(* IEC 61131-3 sources: daoli-st-library/DL_MathData (part 20) *)

(* ---- FC_DL_PeriodJitterCalc.st ---- *)
(*
  Name        : FC_DL_PeriodJitterCalc
  Category    : DL_MathData
  Version     : 1.0.0
  Purpose     : 周期序列抖动统计（双精度数组）：均值、样本标准差（n-1 分母）、峰峰抖动（max-min）；/ Period-sequence jitter statistics over a double-precision array: mean, sample standard deviation (n-1) and peak-to-peak jitter (max-min)
  溯源        : 借 t2-1-lgf-math 的分类/参数域组织，clean-room 实现
  Boundary    : ① 计数域钳位：nCount 钳 0..64（容量常量），少于 2 个有效样本时 bValid = FALSE（样本标准差无定义），返回 0.0 哨兵；
                ② 入口有限性闸：任一被统计元素 NaN（x = x 自反）或 Inf（(x-x) = (x-x) 差判）→ 整体 bValid = FALSE（不静默跳过，防抖动被低估）；
                ③ 除零前置：均值除子为常量 1000 换算与 nCount（>= 2 已闸），标准差除子 nCount-1（>= 1 已闸）；
                ④ 数组下标游标 1..nCount 有界遍历（下标全量钳位），不越容量域；
                ⑤ 返回值 = 峰峰抖动 [s]，bValid = FALSE 时不得使用返回值（上层契约）。
*)
FUNCTION FC_DL_PeriodJitterCalc : LREAL
VAR_INPUT
    afPeriods : ARRAY[1..64] OF LREAL;       (* 周期样本数组（连续周期测量值）[s] / Period samples array *)
    nCount    : INT;                         (* 有效样本数，域 0..64（越域钳位）[个] / Valid sample count, clamped *)
END_VAR
VAR_OUTPUT
    fMean     : LREAL;                       (* 周期均值 [s] / Mean period *)
    fStdDev   : LREAL;                       (* 样本标准差（n-1 分母）[s] / Sample standard deviation *)
    bValid    : BOOL;                        (* 结果有效标志（FALSE 时返回值为哨兵零点）[-] / Result validity flag *)
END_VAR
VAR CONSTANT
    DL_PJC_NMAX  : INT   := 64;              (* 数组容量上限（与形参数组域一致）[个] / Array capacity *)
    DL_PJC_NMIN  : INT   := 2;               (* 样本数下限（标准差最少两点）[个] / Sample lower bound *)
    DL_PJC_EPS   : LREAL := 1.0E-12;         (* 双精度判零容差 [s] / Double-precision epsilon *)
    DL_PJC_ONE   : LREAL := 1.0;             (* 游标递进常量 [-] / Cursor step constant *)
END_VAR
VAR
    _nEff  : INT;                            (* 钳位后生效样本数 [个] / Effective sample count *)
    _nIdx  : INT;                            (* 统计游标（每趟重置，R227）[-] / Stats cursor *)
    _fSum  : LREAL;                          (* Σx 中间量 [s] / Sum intermediate *)
    _fMeanI: LREAL;                          (* 均值中间量 [s] / Mean intermediate *)
    _fVar  : LREAL;                          (* Σ(x-x̄)² 中间量 [s²] / Squared-deviation sum *)
    _fStdI : LREAL;                          (* 标准差中间量 [s] / Std intermediate *)
    _fMin  : LREAL;                          (* 样本最小值 [s] / Sample minimum *)
    _fMax  : LREAL;                          (* 样本最大值 [s] / Sample maximum *)
    _bFin  : BOOL;                           (* 全体样本有限性当拍量 / Joint sample finiteness *)
END_VAR

(* —— 段 0：计数域钳位 + 有限性预置 —— *)
bValid := TRUE;                                                                (* 有效标志预置（任一闸命中即翻 FALSE） / Validity preset *)
_nEff := nCount;                                                               (* 生效样本数初值 / Effective count init *)
IF _nEff < 0 THEN
    _nEff := 0;                                                                (* 计数下限钳 0 / Lower clamp *)
END_IF
IF _nEff > DL_PJC_NMAX THEN
    _nEff := DL_PJC_NMAX;                                                      (* 计数上限钳容量（下标全量钳位） / Upper clamp to capacity *)
END_IF

(* —— 段 1：样本数下限闸（少于 2 点标准差无定义，边界①） —— *)
IF _nEff < DL_PJC_NMIN THEN
    bValid := FALSE;                                                           (* 样本不足：整体无效 / Insufficient samples *)
END_IF

(* —— 段 2：入口有限性闸（逐元素 NaN 自反 + Inf 差判，任一非有限整体拒判，边界②） —— *)
IF bValid THEN
    _bFin := TRUE;                                                             (* 有限性联合量预置 / Finiteness preset *)
    _nIdx := 1;                                                                (* 游标起头 / Cursor reset *)
    WHILE _nIdx <= _nEff DO
        IF NOT ((afPeriods[_nIdx] = afPeriods[_nIdx])                          (* NaN 自反闸 / NaN reflex gate *)
                AND ((afPeriods[_nIdx] - afPeriods[_nIdx]) = (afPeriods[_nIdx] - afPeriods[_nIdx]))) THEN
            _bFin := FALSE;                                                    (* 命中非有限样本 / Non-finite sample hit *)
        END_IF
        _nIdx := _nIdx + DL_PJC_ONE;                                           (* 游标递进（有界遍历） / Cursor advance *)
    END_WHILE
    IF NOT _bFin THEN
        bValid := FALSE;                                                       (* 整体无效（不静默跳过） / Overall invalid *)
    END_IF
END_IF

(* —— 段 3：无效输入早退（出口归零 + 哨兵零点返回） —— *)
IF NOT bValid THEN
    fMean := 0.0;                                                              (* 清均值出口 / Clear mean outlet *)
    fStdDev := 0.0;                                                            (* 清标准差出口 / Clear std outlet *)
    FC_DL_PeriodJitterCalc := 0.0;                                             (* 哨兵零点返回 / Sentinel zero return *)
    RETURN;
END_IF

(* —— 段 4：一趟求 Σx/min/max —— *)
_fSum := 0.0;                                                                  (* Σx 预清 / Sum preset *)
_fMin := afPeriods[1];                                                         (* 最小值初值取首样本 / Min init *)
_fMax := afPeriods[1];                                                         (* 最大值初值取首样本 / Max init *)
_nIdx := 1;                                                                    (* 游标起头（R227） / Cursor reset *)
WHILE _nIdx <= _nEff DO
    _fSum := _fSum + afPeriods[_nIdx];                                         (* Σx [s] / Sum *)
    IF afPeriods[_nIdx] < _fMin THEN
        _fMin := afPeriods[_nIdx];                                             (* 更新最小值 / Update min *)
    END_IF
    IF afPeriods[_nIdx] > _fMax THEN
        _fMax := afPeriods[_nIdx];                                             (* 更新最大值 / Update max *)
    END_IF
    _nIdx := _nIdx + DL_PJC_ONE;                                               (* 游标递进 / Cursor advance *)
END_WHILE

(* —— 段 5：均值与标准差（除子均已过闸，边界③） —— *)
_fMeanI := _fSum / INT_TO_LREAL(_nEff);                                        (* 均值：除子 nEff >= 2 [s] / Mean, divisor >= 2 *)
fMean := _fMeanI;                                                              (* 均值出口 / Mean outlet *)
_fVar := 0.0;                                                                  (* 平方和预清 / Squares preset *)
_nIdx := 1;                                                                    (* 游标重起 / Cursor reset *)
WHILE _nIdx <= _nEff DO
    _fVar := _fVar + (afPeriods[_nIdx] - _fMeanI) * (afPeriods[_nIdx] - _fMeanI);   (* 平方项恒非负 [s²] / Squared deviation *)
    _nIdx := _nIdx + DL_PJC_ONE;                                               (* 游标递进 / Cursor advance *)
END_WHILE
_fStdI := SQRT(_fVar / INT_TO_LREAL(_nEff - 1));                               (* 样本标准差：除子 nEff-1 >= 1 [s] / Sample std, divisor >= 1 *)
fStdDev := _fStdI;                                                             (* 标准差出口 / Std outlet *)

(* —— 段 6：返回峰峰抖动（max-min，无除法） —— *)
FC_DL_PeriodJitterCalc := _fMax - _fMin;                                       (* 峰峰抖动返回 [s] / Peak-to-peak jitter return *)
END_FUNCTION

(* ---- FC_DL_PipeFrictionLoss.st ---- *)
// =====================================================================
// FC_DL_PipeFrictionLoss.st
// Darcy-Weisbach 管道压降纯函数（层流/过渡/湍流自动判别）
// Darcy-Weisbach pipe pressure drop pure function
// 码位: 16#0001_0485 ~ 16#0001_0489 (本件独占 5 槽)
// 修改记录: R29 初版 (按 DISPATCH_R29 序 3)
// =====================================================================
FUNCTION FC_DL_PipeFrictionLoss : BOOL
VAR_INPUT
    bEnable      : BOOL  := TRUE;       // 使能 / Enable
    fFlow_m3h    : REAL  := 0.0;        // 体积流量 ≥0 m³/h / Volumetric flow [m3/h]
    fDia_mm      : REAL  := 50.0;       // 内径 >0 mm / Inner diameter [mm]
    fLen_m       : REAL  := 10.0;       // 直管长度 ≥0 m / Straight length [m]
    fRough_mm    : REAL  := 0.05;       // 绝对粗糙度 ≥0 mm（不锈钢 0.05）/ Absolute roughness [mm]
    fRho_kgm3    : REAL  := 1000.0;     // 密度 >0 kg/m³ / Density [kg/m3]
    fMu_cP       : REAL  := 1.0;        // 动力粘度 >0 cP（水 20℃ 约 1.0）/ Dynamic viscosity [cP]
    fKMinor      : REAL  := 0.0;        // 局部阻力系数和 ≥0 / Minor loss coefficient sum [-]
    fDpMax_kPa   : REAL  := 1000.0;     // 压降量程上限 >0 kPa / Pressure drop full scale [kPa]
    fReLam       : REAL  := 2300.0;     // 层流临界雷诺数 / Laminar critical Re [-]
    fReTurb      : REAL  := 4000.0;     // 湍流起始雷诺数 / Turbulent onset Re [-]
END_VAR
VAR_OUTPUT
    fVel_ms      : REAL;                // 流速 m/s / Velocity [m/s]
    fRe          : REAL;                // 雷诺数 / Reynolds number [-]
    fLambda      : REAL;                // 沿程阻力系数 / Friction factor [-]
    fDp_kPa      : REAL;                // 总压降 kPa / Total pressure drop [kPa]
    bTransition  : BOOL;                // 处于过渡区 / In transition zone
    eErr         : UDINT;               // 错误码 / Error code
END_VAR
VAR
    fArea_m2     : REAL;                // 管道截面积 / Pipe cross-section area [m2]
    fVelSq       : REAL;                // 流速平方 / Velocity squared [(m/s)2]
    fReSafe      : REAL;                // 钳位后安全雷诺数 / Clamped safe Reynolds number [-]
    fLogArg      : REAL;                // log10 参数（钳下限 1E-6）/ log10 argument, clamped [-]
    fLog10Val    : REAL;                // log10 结果 / log10 value [-]
    fDpMaxSafe   : REAL;                // 兜底后量程上限 / Sanitized full scale [kPa]
    fLenSafe     : REAL;                // 长度处理值 / Sanitized length [m]
    bLenNeg      : BOOL;                // 长度负值标记 / Negative length flag
    bClamped     : BOOL;                // 压降钳制标记 / Drop clamped flag
    fDia_m       : REAL;                // 内径转米 / Diameter in meters [m]
    fMu_Pas      : REAL;                // 粘度转 Pa·s / Viscosity in Pa.s [Pa.s]
    fRePow       : REAL;                // Re^0.9 中间量 / Re^0.9 intermediate [-]
    fDpPct       : REAL;                // 直管+局部阻力总系数 / Total resistance factor [-]
END_VAR

// ---------------------------------------------------------------------
// 代码位表（本件独占，勿复用）:
//   16#0001_0485 信息 正常计算完成
//   16#0001_0486 故障 fDia_mm ≤ 0 / fMu_cP ≤ 0 / fRho_kgm3 ≤ 0，或任一输入非有限
//   16#0001_0487 故障 fReLam ≤ 0 / fReTurb ≤ fReLam / fRough_mm < 0 / fKMinor < 0（组态错）
//   16#0001_0488 信息 过渡区（fReLam ≤ Re ≤ fReTurb）→ 按湍流式 + bTransition=TRUE；或压降超上限已钳制
//   16#0001_0489 信息 零流量（fFlow_m3h ≤ 0）→ 三项输出 0、bTransition=FALSE
// ---------------------------------------------------------------------

// 默认输出清零 / Default outputs cleared
fVel_ms     := 0.0;      // 流速清零 / Reset velocity
fRe         := 0.0;      // 雷诺数清零 / Reset Reynolds
fLambda     := 0.0;      // 阻力系数清零 / Reset lambda
fDp_kPa     := 0.0;      // 压降清零 / Reset pressure drop
bTransition := FALSE;    // 过渡区标志复位 / Reset transition flag
eErr        := 16#0001_0485;  // 预置正常码 / Preset normal code

IF NOT bEnable THEN
    // 使能关闭：输出保持 0，不置故障 / Disabled: outputs zero, no fault
    RETURN;   // 直接返回 / Return
END_IF

// ---- 非有限闸 / Finite guard ----
IF (fFlow_m3h <> fFlow_m3h) OR (ABS(fFlow_m3h) >= 1.0E12)
   OR (fDia_mm <> fDia_mm) OR (ABS(fDia_mm) >= 1.0E12)
   OR (fLen_m <> fLen_m) OR (ABS(fLen_m) >= 1.0E12)
   OR (fRough_mm <> fRough_mm) OR (ABS(fRough_mm) >= 1.0E12)
   OR (fRho_kgm3 <> fRho_kgm3) OR (ABS(fRho_kgm3) >= 1.0E12)
   OR (fMu_cP <> fMu_cP) OR (ABS(fMu_cP) >= 1.0E12)
   OR (fKMinor <> fKMinor) OR (ABS(fKMinor) >= 1.0E12)
   OR (fDpMax_kPa <> fDpMax_kPa) OR (ABS(fDpMax_kPa) >= 1.0E12)
   OR (fReLam <> fReLam) OR (ABS(fReLam) >= 1.0E12)
   OR (fReTurb <> fReTurb) OR (ABS(fReTurb) >= 1.0E12) THEN
    eErr := 16#0001_0486;  // 故障：非有限输入 / Fault: non-finite input
    RETURN;                // 输出保持 0 / Outputs stay zero
END_IF

// ---- 物性组态错闸 / Physical property configuration fault ----
IF (fDia_mm <= 0.0) OR (fMu_cP <= 0.0) OR (fRho_kgm3 <= 0.0) THEN
    eErr := 16#0001_0486;  // 故障：径/粘/密非法 / Fault: invalid dia/mu/rho
    RETURN;                // 三输出保持 0，不得抛除零 / Outputs stay zero
END_IF

// ---- 流域组态错闸 / Flow regime configuration fault ----
IF (fReLam <= 0.0) OR (fReTurb <= fReLam)
   OR (fRough_mm < 0.0) OR (fKMinor < 0.0) THEN
    eErr := 16#0001_0487;  // 故障：临界雷诺/粗糙度/局部系数非法 / Fault: invalid regime config
    RETURN;                // 输出保持 0 / Outputs stay zero
END_IF

// ---- 长度负值按 0 处理并置槽 3 / Negative length treated as zero with slot 3 ----
fLenSafe := fLen_m;        // 先原样采用 / Adopt as-is
bLenNeg  := FALSE;         // 标记复位 / Reset flag
IF fLen_m < 0.0 THEN
    fLenSafe := 0.0;       // 按 0 处理 / Treat as zero
    bLenNeg  := TRUE;      // 记录标记 / Mark flag
END_IF

// ---- 量程上限兜底（≤0 按 1000.0，不置错）/ Full-scale fallback ----
IF fDpMax_kPa <= 0.0 THEN
    fDpMaxSafe := 1000.0;  // 兜底 1000 kPa / Fallback 1000 kPa
ELSE
    fDpMaxSafe := fDpMax_kPa;  // 原值 / As-is
END_IF

// ---- 零流量短路路径 / Zero-flow short path ----
IF fFlow_m3h <= 0.0 THEN
    fVel_ms     := 0.0;         // 流速 0 / Zero velocity
    fRe         := 0.0;         // 雷诺数 0 / Zero Reynolds
    fLambda     := 0.0;         // 阻力系数 0 / Zero lambda
    fDp_kPa     := 0.0;         // 压降 0 / Zero drop
    bTransition := FALSE;       // 不在过渡区 / Not in transition
    eErr        := 16#0001_0489;  // 信息级：零流量 / Info: zero flow
    RETURN;                     // 直接返回 / Return
END_IF

// ---- 单位换算与流速 / Unit conversion and velocity ----
fDia_m := fDia_mm / 1000.0;              // mm → m / mm to m
fMu_Pas := fMu_cP / 1000.0;              // cP → Pa·s / cP to Pa.s
fArea_m2 := 3.14159265 * fDia_m * fDia_m / 4.0;  // 截面积 π·d²/4 / Cross-section area [m2]
fVel_ms := (fFlow_m3h / 3600.0) / fArea_m2;      // v = Q/(3600·A) / Velocity [m/s]
fVelSq  := fVel_ms * fVel_ms;                    // v² / Velocity squared

// ---- 雷诺数 Re = v·d·ρ/μ / Reynolds number ----
fRe := fVel_ms * fDia_m * fRho_kgm3 / fMu_Pas;   // 雷诺数 / Reynolds number [-]

// ---- Re 钳 1.0 防幂运算溢出（Re=0 时 5.74/Re^0.9 无定义）/ Clamp Re to 1.0 ----
IF fRe < 1.0 THEN
    fReSafe := 1.0;   // 钳下限 / Clamp minimum
ELSE
    fReSafe := fRe;   // 原值 / As-is
END_IF

// ---- 分流域计算 λ / Regime-based lambda ----
bTransition := FALSE;   // 过渡区标志复位 / Reset transition flag
IF fRe < fReLam THEN
    // 层流：λ = 64/Re（ReSafe ≥ 1.0 保证分母安全）/ Laminar
    fLambda := 64.0 / fReSafe;               // 层流阻力系数 / Laminar friction factor
ELSIF fRe <= fReTurb THEN
    // 过渡区：按湍流式算 + 信息级（不中断）/ Transition: turbulent formula + info
    bTransition := TRUE;                     // 标记过渡区 / Mark transition
    eErr        := 16#0001_0488;             // 信息级：过渡区 / Info: transition
    fRePow := EXPT(fReSafe, 0.9);            // Re^0.9 / Re to power 0.9
    fLogArg := (fRough_mm / (3.7 * fDia_mm)) + (5.74 / fRePow);  // Swamee-Jain 内项 / SJ argument
    IF fLogArg < 1.0E-6 THEN
        fLogArg := 1.0E-6;                   // 钳下限防 log10 奇点 / Clamp to avoid singularity
    END_IF
    fLog10Val := LOG(fLogArg) / 2.302585093; // 自然对数换底 log10 / Convert to log10
    IF ABS(fLog10Val) < 1.0E-9 THEN
        fLog10Val := 1.0E-9;                 // 防平方后除零 / Guard division
    END_IF
    fLambda := 0.25 / (fLog10Val * fLog10Val);  // 湍流式 λ / Turbulent friction factor
ELSE
    // 湍流：Swamee-Jain 显式式 / Turbulent: Swamee-Jain explicit
    fRePow := EXPT(fReSafe, 0.9);            // Re^0.9 / Re to power 0.9
    fLogArg := (fRough_mm / (3.7 * fDia_mm)) + (5.74 / fRePow);  // 内项 / SJ argument
    IF fLogArg < 1.0E-6 THEN
        fLogArg := 1.0E-6;                   // 钳下限 / Clamp minimum
    END_IF
    fLog10Val := LOG(fLogArg) / 2.302585093; // 换底 log10 / Convert to log10
    IF ABS(fLog10Val) < 1.0E-9 THEN
        fLog10Val := 1.0E-9;                 // 防除零 / Guard division
    END_IF
    fLambda := 0.25 / (fLog10Val * fLog10Val);  // λ / Friction factor
END_IF

// ---- 总压降 Δp = (λ·L/d + ΣK)·ρ·v²/2 / Total pressure drop ----
fDpPct := (fLambda * fLenSafe / fDia_m) + fKMinor;  // 总阻力系数 / Total resistance factor
fDp_kPa := (fDpPct * fRho_kgm3 * fVelSq / 2.0) / 1000.0;  // Pa → kPa / Pressure drop [kPa]

// ---- 量程钳制（信息级）/ Full-scale clamp (info level) ----
bClamped := FALSE;               // 钳制标记复位 / Reset clamp flag
IF fDp_kPa > fDpMaxSafe THEN
    fDp_kPa  := fDpMaxSafe;      // 钳到上限 / Clamp to full scale
    bClamped := TRUE;            // 记录钳制 / Mark clamped
END_IF

// ---- 信息级汇总：长度负值/钳制覆盖正常码 / Info aggregation ----
IF bLenNeg OR bClamped THEN
    eErr := 16#0001_0488;        // 信息：过渡区或钳制共用槽 4 / Info: transition or clamp slot
END_IF

// 正常完成，返回 TRUE / Normal completion
FC_DL_PipeFrictionLoss := TRUE;  // 函数返回值 / Function result

END_FUNCTION

(* ---- FC_DL_PlasmaPowerDensityCalc.st ---- *)
(*
  DL Factory R88 | FC_DL_PlasmaPowerDensityCalc
  功能：算等离子体功率密度 P/A，并按 1~5 W/cm² 工艺带宽判合格
  开源溯源：无（clean-room 自研，依据公开工艺公式 功率密度定义式 P/A，许可证=MIT，借鉴点=公式结构）
  规则：R1-R16 全遵守；R88 简单件标量形（纯标量入参出参，无循环体、无方法、无属性、无数组）
*)
FUNCTION FC_DL_PlasmaPowerDensityCalc : REAL
VAR_INPUT
    fPowerW : REAL := 800.0; // 射频/直流输入功率 P [W] / RF or DC input power [W]
    fAreaCm2 : REAL := 400.0; // 电极（或基片）有效面积 A [cm²] / effective electrode area [cm^2]
    fMinWPerCm2 : REAL := 1.0; // 功率密度允许下限 [W/cm²] / lower density band [W/cm^2]
    fMaxWPerCm2 : REAL := 5.0; // 功率密度允许上限 [W/cm²] / upper density band [W/cm^2]
END_VAR
VAR_OUTPUT
    fDensityWPerCm2 : REAL; // 功率密度 [W/cm²] / power density [W/cm^2]
    xInBand : BOOL; // TRUE=功率密度落在允许带宽内 [-] / TRUE when inside the band [-]
END_VAR
VAR
    fAreaDenom : REAL; // 面积分母（除零判据） [cm²] / area divisor [cm^2]
END_VAR

// 段 1｜出口预置
FC_DL_PlasmaPowerDensityCalc := -1.0; // 哨兵返回 -1（无效） [-] / sentinel return -1, invalid [-]
fDensityWPerCm2 := 0.0; // 功率密度预置零 [W/cm²] / density preset zero [W/cm^2]
xInBand := FALSE; // 带宽位预置 FALSE（未判定前不认合格） [-] / band flag preset false [-]
fAreaDenom := 0.0; // 面积分母预置零 [cm²] / area divisor preset zero [cm^2]

// 段 2｜非有限拦截 + 域闸
IF NOT (fPowerW > -1.0E30 AND fPowerW < 1.0E30) OR NOT (fAreaCm2 > -1.0E30 AND fAreaCm2 < 1.0E30) THEN
    RETURN; // 功率/面积任一非有限即拒算 [-] / any non finite input rejected [-]
END_IF
IF NOT (fMinWPerCm2 > -1.0E30 AND fMinWPerCm2 < 1.0E30) OR NOT (fMaxWPerCm2 > -1.0E30 AND fMaxWPerCm2 < 1.0E30) THEN
    RETURN; // 带宽上下限任一非有限则判据静默失效，故先拦 [W/cm²] / band limits must be finite [W/cm^2]
END_IF
IF fPowerW < 0.0 THEN
    RETURN; // 功率非负闸（负功率无物理意义） [W] / non negative power gate [W]
END_IF
IF fAreaCm2 < 1.0E-9 THEN
    RETURN; // 面积正域闸（同时是分母，防除零） [cm²] / positive area, also the divisor [cm^2]
END_IF
IF fMinWPerCm2 <= 0.0 OR fMaxWPerCm2 <= fMinWPerCm2 THEN
    RETURN; // 带宽自洽闸：下限须为正、上限须严格大于下限 [W/cm²] / band consistency gate [W/cm^2]
END_IF

// 段 3｜计算
fAreaDenom := fAreaCm2; // 取面积作除数 [cm²] / take the area as divisor [cm^2]
IF fAreaDenom < 1.0E-9 THEN
    RETURN; // 除法前分母闸：面积必须大于 1E-9 才可作除数 [cm²] / denominator gate before the division [cm^2]
END_IF
fDensityWPerCm2 := fPowerW / fAreaDenom; // W ÷ cm² = W/cm²，功率密度 [W/cm²] / [W] / [cm^2] = [W/cm^2]

// 段 4｜判定与饱和
IF NOT (fDensityWPerCm2 > -1.0E30 AND fDensityWPerCm2 < 1.0E30) THEN
    RETURN; // 结果非有限再拦一次 [-] / re-check the result for finiteness [-]
END_IF
xInBand := (fDensityWPerCm2 >= fMinWPerCm2) AND (fDensityWPerCm2 <= fMaxWPerCm2); // 双侧闭区间直比 [W/cm²] / closed two sided band compare [W/cm^2]

// 段 5｜出口自检
IF fDensityWPerCm2 < 0.0 THEN
    RETURN; // 出口自检：功率密度不得为负（负值说明输入符号错） [W/cm²] / must not be negative [W/cm^2]
END_IF
FC_DL_PlasmaPowerDensityCalc := fDensityWPerCm2; // 返回功率密度 [W/cm²] / return the power density [W/cm^2]
END_FUNCTION

(* ---- FC_DL_PolarDecomp2D.st ---- *)
(*==============================================================================
 * 组件名称 (Component)  : FC_DL_PolarDecomp2D
 * 所属子库 (Sublibrary) : DL_MathData
 * 当前版本 (Version)    : 1.0.0
 * 兼容性 (Platform)     : CODESYS 3.5+ / TwinCAT 3 / 汇川 InoProShop / 施耐德 Machine Expert
 *                         仅依赖 Standard.library（SQRT / ATAN / ABS），零厂商私有库
 * 功能描述 (Function)   : 2D 矩阵极分解（纯函数 FC）。对 2×2 矩阵 M 求
 *                         M = R·S：S = (MᵀM)^(1/2) 对称正定部分，R 旋转部分；
 *                         输出主方向角 θ（S 的最大特征向量角）与两个奇异值
 *                         σ1 >= σ2（谱半径语义）。算法：MᵀM 的对称表示
 *                         [a b; b c]，特征值 λ = (T ± √(D²+4b²))/2（T=a+c,
 *                         D=a-c），θ = 0.5·atan2(2b, a-c)。与 Matrix3Inverse
 *                         （求逆）/Affine2D*（仿射组合）分工：谱语义首次入库。
 * 来源标签 (Origin)     : 源矩阵 T2-1 LGF Math ◐ 待挖子项（R25 备注既有），自研 clean-room
 * 边界语义 (Boundary)   : ① 输入 NaN/Inf → 返回 FALSE，输出哨兵 0（还原方向
 *                         不饱和、哨兵 + 有效性位，R81）；
 *                         ② 零矩阵（λ1 <= eps）→ 返回 FALSE（主方向无定义）；
 *                         ③ atan2 本地实现（纯 ATAN 四象限组装），贴轴归属
 *                         写死：y = 0 且 x < 0 归 y >= 0 支，值域 (-π, π]（R52）；
 *                         ④ 除法仅出现在 atan2 域内（x ≠ 0 分支），无除零。
 * 输出语义 (Fallback)   : 返回 FALSE → fTheta/fSigma1/fSigma2 哨兵 0（调用方
 *                         以返回值判有效性，非故障级）。
 * 码位     (Codes)      : 按 R297 范式零 16# 码位硬编码（纯函数无错误码）。
 * 红线自检 (Redline)    : 7 项红线已自检：R1 零全局 ✓｜R2 零物理地址 ✓｜R3 纯 IEC ✓
 *                         R4 除零（atan2 分支闸）/NaN 哨兵 ✓｜R5 双语同行注释 ✓
 *                         R6 纯函数无顺序逻辑（CASE 无涉）✓｜R7 无定时器实例 ✓
 * 验收向量 (Acceptance) : V1 M=diag(2,1) → σ1=2.0、σ2=1.0、θ=0.0（对角阵
 *                         主方向沿 x 轴）；
 *                         V2 纯旋转 45°（MᵀM=I）→ σ1=σ2=1.0、θ=0.0（各向
 *                         同性退化，θ 无定义取 0 并在头注释声明）；
 *                         V3 剪切 [[1,1],[0,1]] → σ1=1.618034（黄金比）、
 *                         σ2=0.618034、θ≈1.0172 rad（公开数值可复算）。
 * 修订历史 (Revision)   : 2026-11-20  v1.0.0  R51 首版（批 3 · 序号 15）
 *==============================================================================*)
FUNCTION FC_DL_PolarDecomp2D : BOOL     // 返回 TRUE = 分解有效（θ/σ 可信）/ TRUE = decomposition valid
VAR_INPUT
    fM11 : LREAL;                        (* 矩阵 M 第 1 行第 1 列 [-] / Matrix element m11 *)
    fM12 : LREAL;                        (* 矩阵 M 第 1 行第 2 列 [-] / Matrix element m12 *)
    fM21 : LREAL;                        (* 矩阵 M 第 2 行第 1 列 [-] / Matrix element m21 *)
    fM22 : LREAL;                        (* 矩阵 M 第 2 行第 2 列 [-] / Matrix element m22 *)
END_VAR
VAR_OUTPUT
    fTheta  : LREAL;                     (* 主方向角（S 最大特征向量角）[rad] / Principal direction angle *)
    fSigma1 : LREAL;                     (* 奇异值 1（σ1 >= σ2）[-] / Largest singular value *)
    fSigma2 : LREAL;                     (* 奇异值 2 [-] / Smaller singular value *)
END_VAR
VAR
    fA    : LREAL;                       (* MᵀM 对称元素 a = m11²+m21² [-] / Symmetric element a *)
    fB    : LREAL;                       (* MᵀM 对称元素 b = m11·m12+m21·m22 [-] / Symmetric element b *)
    fC    : LREAL;                       (* MᵀM 对称元素 c = m12²+m22² [-] / Symmetric element c *)
    fT    : LREAL;                       (* 迹 T = a + c [-] / Trace *)
    fD    : LREAL;                       (* 对角差 D = a - c [-] / Diagonal difference *)
    fDisc : LREAL;                       (* 判别式 D² + 4b² [-] / Discriminant *)
    fL1   : LREAL;                       (* 特征值 λ1 = (T+√disc)/2 [-] / Eigenvalue 1 *)
    fL2   : LREAL;                       (* 特征值 λ2 = (T-√disc)/2 [-] / Eigenvalue 2 *)
    fAx   : LREAL;                       (* atan2 实参 x = a - c [-] / atan2 argument x *)
    fAy   : LREAL;                       (* atan2 实参 y = 2b [-] / atan2 argument y *)
    fAng  : LREAL;                       (* atan2 结果工作量 [rad] / atan2 result work *)
END_VAR
VAR CONSTANT
    DL_PDC_EPS : LREAL := 1.0E-12;       (* 特征值判零容差 [-] / Eigenvalue epsilon *)
    DL_PDC_PI  : LREAL := 3.14159265358979324;   (* π（LREAL 精度字面量，R51①）[rad] / Pi *)
    DL_PDC_PI2 : LREAL := 1.57079632679489662;   (* π/2 [rad] / Half pi *)
END_VAR

(* —— 段 0：输出哨兵预置（还原方向不饱和，R81） —— *)
fTheta := 0.0;                           (* θ 哨兵 0 / Theta sentinel *)
fSigma1 := 0.0;                          (* σ1 哨兵 0 / Sigma1 sentinel *)
fSigma2 := 0.0;                          (* σ2 哨兵 0 / Sigma2 sentinel *)
FC_DL_PolarDecomp2D := FALSE;            (* 返回值预置无效 / Return preset invalid *)

(* —— 段 1：输入非有限闸（NaN 自反 + Inf 差判，R79） —— *)
IF (fM11 <> fM11) OR ((fM11 - fM11) <> (fM11 - fM11))
   OR (fM12 <> fM12) OR ((fM12 - fM12) <> (fM12 - fM12))
   OR (fM21 <> fM21) OR ((fM21 - fM21) <> (fM21 - fM21))
   OR (fM22 <> fM22) OR ((fM22 - fM22) <> (fM22 - fM22)) THEN
    RETURN;                              (* 非有限输入：哨兵 + FALSE 早退（变换集合 = 哨兵全零，无后处理须补，R94） / Non-finite: early return with sentinels *)
END_IF

(* —— 段 2：MᵀM 对称表示与特征分解 —— *)
fA := fM11 * fM11 + fM21 * fM21;         (* a = m11² + m21² / Element a *)
fB := fM11 * fM12 + fM21 * fM22;         (* b = m11·m12 + m21·m22 / Element b *)
fC := fM12 * fM12 + fM22 * fM22;         (* c = m12² + m22² / Element c *)
fT := fA + fC;                           (* 迹 / Trace *)
fD := fA - fC;                           (* 对角差 / Diagonal diff *)
fDisc := fD * fD + 4.0 * fB * fB;        (* 判别式（≥ 0 结构性成立，MᵀM 半正定） / Discriminant *)
fL1 := 0.5 * (fT + SQRT(fDisc));         (* λ1（SQRT 实参 ≥ 0 无域违例） / Eigenvalue 1 *)
fL2 := 0.5 * (fT - SQRT(fDisc));         (* λ2 / Eigenvalue 2 *)
IF fL1 <= DL_PDC_EPS THEN
    RETURN;                              (* 零矩阵：主方向无定义，哨兵 + FALSE（边界②） / Zero matrix: return FALSE *)
END_IF

(* —— 段 3：本地 atan2 四象限组装（贴轴归属写死：y=0 且 x<0 归 y>=0 支，值域 (-π, π]，R52） —— *)
fAx := fA - fC;                          (* 实参 x / Argument x *)
fAy := 2.0 * fB;                         (* 实参 y / Argument y *)
IF fAx > 0.0 THEN
    fAng := ATAN(fAy / fAx);             (* 右半平面：除子 x > 0 无除零 / Right half: divide gated *)
ELSIF fAx < 0.0 THEN
    IF fAy >= 0.0 THEN
        fAng := ATAN(fAy / fAx) + DL_PDC_PI;   (* 上左半平面（含贴轴 y=0,x<0 → π） / Upper-left incl. axis rule *)
    ELSE
        fAng := ATAN(fAy / fAx) - DL_PDC_PI;   (* 下左半平面 / Lower-left *)
    END_IF
ELSE                                     (* x = 0 贴轴支 / Axis branch *)
    IF fAy > 0.0 THEN
        fAng := DL_PDC_PI2;              (* +π/2 / +pi/2 *)
    ELSIF fAy < 0.0 THEN
        fAng := -DL_PDC_PI2;             (* -π/2 / -pi/2 *)
    ELSE
        fAng := 0.0;                     (* x=y=0：退化方向取 0（各向同性，与 V2 声明一致） / Degenerate: zero *)
    END_IF
END_IF

(* —— 段 4：输出映射（σ 由 λ 开方，λ >= 0 结构性保证无域违例） —— *)
fTheta := 0.5 * fAng;                    (* 主方向角 = 半角（特征向量角公式） / Principal angle *)
fSigma1 := SQRT(fL1);                    (* σ1 = √λ1（λ1 > eps 已闸） / Sigma1 *)
fSigma2 := SQRT(fL2);                    (* σ2 = √λ2（λ2 >= 0 半正定） / Sigma2 *)
FC_DL_PolarDecomp2D := TRUE;             (* 分解有效 / Valid *)
END_FUNCTION

(* ---- FC_DL_PolyEvalHorner.st ---- *)
(*
    组件名称 : FC_DL_PolyEvalHorner
    所属子库 : DL_MathData
    当前版本 : 1.0.0
    兼 容 性 : CODESYS V3.5+ / TwinCAT 3 / 汇川 InoProShop；仅依赖 Standard.library
    功能描述 : Horner 法多项式求值内核，PT100 Callendar-Van Dusen、热电偶 NIST 多项式、传感器多点拟合的公共出口。
              取舍 ①：升幂系数 a0..an + Horner 递推，n 次乘加内完成求值；相比「逐项 x^i × a_i」少一半乘法、
              少 n 次幂运算，更重要的是不产生中间大数（x^i 在高阶处会先溢出，再乘 a_i 又变回来，纯损失精度）。
              取舍 ②：前导零系数自动降阶 —— 上位机配置表常把 4 阶多项式填进 8 阶槽位，尾部全是 0.0；
              不降阶就会白做 4 次「乘 0 加 0」，把尾数误差放大并拖慢扫描。降阶后 nEffOrder 一并出口，
              调用方能看到「实际用了几阶」。
              取舍 ③：系数用 VAR_IN_OUT 免拷贝 —— 8 阶 LREAL 数组按值传参在部分平台是一次整段复制，
              本件是高频调用内核算术路径，不能付这个代价。
              取舍 ④：中间量逐阶判非有限 —— 溢出可能发生在中途而终值又被后续系数拉回有限域，
              只查终值会漏掉「中间已脏、结果恰好像样」的假值。
    开源溯源 : 原创实现。与存量 FC_DL_MultiPointLinear / FC_DL_InterpolateTable2D 的边界：那两件是分段线性/双线性，；本件为 IEC 61131-3 标准语义的道莅防御性实现（原创实现，零外部源码复制）。
              本件是单一多项式。无外部源码参考，码位与分级 100% 自有。
    本文件内含 : FUNCTION FC_DL_PolyEvalHorner（单 POU，无配套类型）
    依 赖 : 无 DL_ 内部依赖；Standard.library: 无
    红线自检 : R1 ✓ 零全局变量与外部变量 ｜ R2 ✓ 零物理 IO 地址
              R3 ✓ 纯 IEC 61131-3 ｜ R4 ✓ 阶数闸 + 非有限闸 + WHILE 守卫计数器 + 中间量逐阶复检
              R5 ✓ 全变量中英双语同行注释 ｜ R6 N/A 纯函数无顺序状态机，无 CASE 可写
              R7 N/A 无定时器、无沿检测实例 ｜ R8 ✓ 阶数上限、容差、有限域全常量化
    错误码   : 16#0001_043A [信息级] 前导零系数已降阶，nEffOrder < nOrder，bValid = TRUE
               16#0001_043B [信息级] 预留禁用（不得挪用）
               16#0001_0375 [故障级] 阶数越界（< 0 或 > DL_POLY_MAX_ORDER），返回 0，bValid = FALSE
               16#0001_0376 [故障级] fX 或参与运算的系数非有限，返回 0，bValid = FALSE
               16#0001_0377 [故障级] 中间量或结果溢出，返回 0，bValid = FALSE
    码位总账 : 16#0001_043A 用 / 16#0001_043B 预留 ｜ 16#0001_0375 用 / 16#0001_0376 用 / 16#0001_0377 用
    遗留假设 : ① FOR 循环在初值小于终值时（如 nEffOrder = 0 时的 DOWNTO）执行零次，IEC 语义保证；
              本件仍用 IF nEffOrder > 0 显式包一层，不依赖该语义。此写法为双保险，未三平台逐一实测。
              ② 无时间/日期与字符串内建依赖，编译门槛未见风险。
    修订历史 :
        2026-11-16  v1.0.0  首版，R21 批次 1 入库
*)
FUNCTION FC_DL_PolyEvalHorner : LREAL
VAR_INPUT
    nOrder          : INT := 0;                  // 阶数，0~DL_POLY_MAX_ORDER，越界即拒算 [阶] / polynomial order, rejected when out of range [order]
    fX              : LREAL := 0.0;              // 自变量，如温度 [工程单位] / independent variable, e.g. temperature [engineering unit]
END_VAR
VAR_IN_OUT
    afCoeff         : ARRAY[0..DL_POLY_MAX_ORDER] OF LREAL;   // 升幂系数 a0..an，下标即幂次；前导零自动降阶 [系数] / ascending coefficients, the index is the power [coefficient]
END_VAR
VAR_OUTPUT
    eErr            : UDINT;                     // 错误码，0=正常；16#0001_04XX 信息级 / 16#0001_03XX 故障级 / error id, 0=ok
    bError          : BOOL;                      // 故障级标志，eErr 落 16#0001_03XX 时为 TRUE / fault flag, TRUE on fault-level eErr
    bValid          : BOOL;                      // 求值结果是否可用 / evaluation usable flag
    nEffOrder       : INT;                       // 实际使用的阶数（降阶后）[阶] / effective order after the leading zero reduction [order]
END_VAR
VAR
    nEff            : INT;                       // 降阶游标 [阶] / reduction cursor [order]
    nGuard          : DINT;                      // WHILE 防死锁守卫计数 [次] / loop guard counter [count]
    nIdx            : INT;                       // Horner 递推下标 [阶] / Horner recursion index [order]
    nJ              : INT;                       // 升序循环变量（镜像下标用）[阶] / ascending loop var for mirrored index
    fAcc            : LREAL;                     // 累加工作寄存器 [工程单位] / accumulation working register [engineering unit]
    bOverflow       : BOOL;                      // 中间量溢出标志 / intermediate overflow flag
END_VAR
VAR CONSTANT
    DL_POLY_MAX_ORDER   : INT := 8;                            // 最高阶数（PT100 CVD 4 阶、热电偶 NIST ≤ 8 阶）[阶] / highest supported order [order]
    DL_POLY_GUARD_MAX   : DINT := 32;                          // 降阶 WHILE 守卫上限，远大于 8，纯防御 [次] / guard limit for the reduction loop, pure defence [count]
    DL_FLOAT_EPS        : LREAL := 1.0E-12;                    // 判零容差，系数降阶用（禁 = 0 判等）[无量纲] / zero tolerance for the reduction test [dimensionless]
    DL_LREAL_MAX_FINITE : LREAL := 1.7976931348623157E308;     // LREAL 最大有限值 [无量纲] / largest finite LREAL [dimensionless]
    DL_LREAL_ZERO       : LREAL := 0.0;                        // 零哨兵 [无量纲] / zero sentinel [dimensionless]
    DL_INT_ONE          : INT := 1;                            // 单位哨兵，避免裸 1 [无量纲] / unity sentinel [dimensionless]
    DL_ERR_NONE         : UDINT := 16#0000_0000;               // 无故障 / no error
END_VAR

// 段 1｜返回值与错误状态预置 / segment 1, preset the return value and the error state
FC_DL_PolyEvalHorner := DL_LREAL_ZERO;  // 故障缺省返回 0 / fault default returns zero
eErr        := DL_ERR_NONE;             // 预置无错误 / preset no error
bError      := FALSE;                   // 预置无故障 / preset no fault
bValid      := FALSE;                   // 预置结果不可用 / preset unusable
nEffOrder   := 0;                       // 预置实际阶数 0 / preset the effective order to zero
nEff        := 0;                       // 预置降阶游标 / preset the reduction cursor

// 段 2｜阶数闸：越界一律拒算，不做静默钳位 / segment 2, order gate, reject instead of silently clamping
IF (nOrder < 0) OR (nOrder > DL_POLY_MAX_ORDER) THEN
    eErr   := 16#0001_0375;             // 阶数越界（故障级）/ order out of range, fault level
    bError := TRUE;                     // 置故障标志 / raise the fault flag
    RETURN;                             // 返回 0，bValid 保持 FALSE / return zero, bValid stays FALSE
END_IF

// 段 3｜自变量有限性闸 / segment 3, independent variable finiteness gate
IF (fX <> fX) OR (ABS(fX) > DL_LREAL_MAX_FINITE) THEN
    eErr   := 16#0001_0376;             // 自变量非有限（故障级）/ non-finite independent variable, fault level
    bError := TRUE;                     // 置故障标志 / raise the fault flag
    RETURN;                             // 返回 0，bValid 保持 FALSE / return zero, bValid stays FALSE
END_IF

// 段 4｜前导零降阶：WHILE 必带守卫计数器，超限即判故障 / segment 4, leading zero reduction with a guarded WHILE
nEff   := nOrder;                       // 从声明阶数起降 / start from the declared order
nGuard := 0;                            // 守卫计数清零 / clear the guard counter
WHILE (nEff > 0) AND (ABS(afCoeff[nEff]) < DL_FLOAT_EPS) AND (nGuard <= DL_POLY_GUARD_MAX) DO
    nEff   := nEff - 1;                 // 最高阶系数为零，降一阶 / the top coefficient is zero, drop one order
    nGuard := nGuard + 1;               // 守卫递增 / increment the guard
END_WHILE
IF nGuard > DL_POLY_GUARD_MAX THEN
    eErr   := 16#0001_0377;             // 降阶失控判溢出类故障（理论不可达，纯防御）/ reduction runaway, defensive only
    bError := TRUE;                     // 置故障标志 / raise the fault flag
    RETURN;                             // 返回 0 / return zero
END_IF
nEffOrder := nEff;                      // 出口实际阶数 / publish the effective order
IF nEff < nOrder THEN
    eErr := 16#0001_043A;               // 前导零已降阶（信息级，不置 bError）/ leading zeros reduced, info level
END_IF

// 段 5｜参与运算的系数有限性闸：只查 0..nEff，未参与的槽位不参与判据 / segment 5, finiteness of the participating coefficients only
FOR nIdx := 0 TO nEff DO
    IF (afCoeff[nIdx] <> afCoeff[nIdx]) OR (ABS(afCoeff[nIdx]) > DL_LREAL_MAX_FINITE) THEN
        eErr   := 16#0001_0376;         // 系数非有限（故障级）/ non-finite coefficient, fault level
        bError := TRUE;                 // 置故障标志 / raise the fault flag
        RETURN;                         // 返回 0，bValid 保持 FALSE / return zero, bValid stays FALSE
    END_IF
END_FOR

// 段 6｜Horner 递推：nEff 次乘加，逐阶复检中间量 / segment 6, Horner recursion with per-step re-check
fAcc       := afCoeff[nEff];            // 最高阶系数作为起值 / seed with the top coefficient
bOverflow  := FALSE;                    // 溢出标志清零 / clear the overflow flag
IF nEff > 0 THEN
    FOR nJ := 0 TO (nEff - 1) DO
        nIdx := (nEff - 1) - nJ;                                              // 镜像下标：R509 禁 DOWNTO / mirrored index, DOWNTO unsupported
        fAcc := fAcc * fX + afCoeff[nIdx];                                  // 一次乘加降一阶 / one multiply-add per order
        IF (fAcc <> fAcc) OR (ABS(fAcc) > DL_LREAL_MAX_FINITE) THEN          // 中间量非有限即溢出 / a non-finite intermediate means overflow
            bOverflow := TRUE;                                              // 锁定溢出标志 / latch the overflow flag
        END_IF
    END_FOR
END_IF

// 段 7｜出口复检：中间溢出与终值溢出同码 / segment 7, exit re-check, an intermediate or final overflow shares one code
IF bOverflow OR (ABS(fAcc) > DL_LREAL_MAX_FINITE) THEN
    FC_DL_PolyEvalHorner := DL_LREAL_ZERO;  // 溢出不给伪值 / never emit a pseudo value on overflow
    eErr   := 16#0001_0377;                 // 结果溢出（故障级）/ result overflow, fault level
    bError := TRUE;                         // 置故障标志 / raise the fault flag
    RETURN;                                 // bValid 保持 FALSE / bValid stays FALSE
END_IF

// 段 8｜出口 / segment 8, exit
FC_DL_PolyEvalHorner := fAcc;           // 输出求值结果 / publish the evaluation result
bValid := TRUE;                         // 结果可用 / the result is usable
END_FUNCTION

(* ---- FC_DL_PolygonArea.st ---- *)
(*==============================================================================
 * 组件名称 (Component)  : FC_DL_PolygonArea
 * 所属子库 (Sublibrary) : DL_MathData
 * 当前版本 (Version)    : 1.0.0
 * 兼容性   (Platform)   : CODESYS 3.5 / TwinCAT 3 / 汇川 InoProShop / Machine Expert
 *                         仅依赖 Standard.library（ABS / MOD），全 LREAL 运算，无状态
 * 功能描述 (Function)   : 平面多边形有向面积、绝对面积与质心坐标（鞋带公式 / Green 定理的
 *                         离散形式）。用于视觉定位的料框有效面积、零件轮廓面积校验、
 *                         机器人平面抓取中心计算、皮带跑偏区域判断。
 *                         返回值即绝对面积，有向面积符号经 bCcw 输出，供调用方判断轮廓
 *                         绕向（多数视觉库输出顺时针轮廓，需要翻转才能与机器人坐标系一致）。
 *
 * 【失真与语义披露 / Distortion disclosure】
 *   1) 自交多边形：鞋带公式返回的是代数面积（正负抵消），不是几何面积。结果无几何意义，
 *      调用方必须保证输入是简单多边形；视觉轮廓应先按角度排序并去重，再送进来。
 *   2) 顶点约定"末点不重复首点"。若调用方重复传入首点，面积仍正确，但质心会偏移
 *      （重复点参与一次额外的零面积边，却多算了一次顶点权重）。检测办法：首末点距离
 *      小于 eps 时把 nCount 减 1 再调用。
 *   3) 退化（点数 < 3、共线、零面积）时质心返回顶点算术平均，而不是 (0,0)：
 *      (0,0) 会让机器人在异常时朝原点狂奔，算术平均至少落在轮廓附近。
 *   4) 必须用 LREAL：32 点 × 1e6 mm 坐标的叉积累加可达 1e12，REAL 的 24 位尾数在这个
 *      量级已经丢掉 5 位有效数字，面积会算出负偏差。
 *
 * 开源溯源 (Origin)     : 原创实现（参考西门子 LGF 数学功能组中平面几何族的分类位置，
 *                         鞋带公式为公开数学方法，clean-room 独立实现）
 * 依赖     (Depends)    : 无 DL_ 内部依赖；Standard.library: ABS / MOD
 * 红线自检 (Redline)    : R1 ✓ 零全局变量表与外部变量引用 ｜ R2 ✓ 零物理 IO 地址直写
 *                         R3 ✓ 纯 IEC 61131-3（MOD 取模闭合索引，无负索引）
 *                         R4 ✓ 点数双向钳位 + 索引只经 MOD + 面积零容差 + 质心分母判零
 *                         R5 ✓ 全变量中英双语同行注释 ｜ R6 N/A（无状态机）｜ R7 N/A（无实例调用）
 * 修订历史 (Revision)   :
 *   2026-11-14  v1.0.0  首版入库（Phase 1 收口批次 · R3）
 *============================================================================*)
FUNCTION FC_DL_PolygonArea : LREAL
VAR_IN_OUT
    afX : ARRAY[0..31] OF LREAL;          // 顶点 X 序列，末点不重复首点（上限 32 点）/ Vertex X, not closed, max 32
    afY : ARRAY[0..31] OF LREAL;          // 顶点 Y 序列（上限 32 点）/ Vertex Y, max 32
END_VAR
VAR_INPUT
    nCount : INT;                         // 顶点数，合法域 3..32 / Vertex count, valid 3..32
END_VAR
VAR_OUTPUT
    fCentroidX  : LREAL;                  // 质心 X [mm] / Centroid X [mm]
    fCentroidY  : LREAL;                  // 质心 Y [mm] / Centroid Y [mm]
    bCcw        : BOOL;                   // TRUE = 逆时针（右手系）/ TRUE = counter-clockwise, right-handed
    bDegenerate : BOOL;                   // TRUE = 退化（共线或面积为零）/ TRUE = degenerate polygon
    uErrorId    : UDINT;                  // 故障码，0 = 无故障 / Error code, 0 = no error
END_VAR
VAR
    nI      : INT;                        // 顶点索引 / Vertex index
    nJ      : INT;                        // 下一顶点索引 (nI + 1) MOD nCount / Next vertex index
    nCnt    : INT;                        // 钳位后的有效顶点数 / Clamped effective vertex count
    nGuard  : INT;                        // 循环防死锁计数器 / Loop guard counter
    fCross  : LREAL;                      // 单边叉积项 [mm^2] / Per-edge cross term [mm^2]
    fArea2  : LREAL;                      // 二倍有向面积 [mm^2] / Twice the signed area [mm^2]
    fCxAcc  : LREAL;                      // 质心 X 累加 [mm^3] / Centroid X accumulator [mm^3]
    fCyAcc  : LREAL;                      // 质心 Y 累加 [mm^3] / Centroid Y accumulator [mm^3]
    fDen    : LREAL;                      // 质心公式分母 3×fArea2 [mm^2] / Centroid denominator
    fMeanX  : LREAL;                      // 顶点算术平均 X（退化回退）[mm] / Mean X fallback [mm]
    fMeanY  : LREAL;                      // 顶点算术平均 Y（退化回退）[mm] / Mean Y fallback [mm]
END_VAR
VAR CONSTANT
    DL_PGA_PTS_MIN : INT   := 3;          // 最少顶点数 / Minimum vertex count
    DL_PGA_PTS_MAX : INT   := 32;         // 最多顶点数，等于数组维度 / Maximum vertex count, equals the array size
    DL_PGA_EPS     : LREAL := 1.0E-12;    // 面积零判定容差 [mm^2] / Zero-area tolerance [mm^2]
    DL_PGA_TWO     : LREAL := 2.0;        // 面积公式分母常数 / Area denominator constant
    DL_PGA_THREE   : LREAL := 3.0;        // 质心分母常数，6×(A2/2) 折算为 3×A2 / Reduced centroid denominator
END_VAR

(*------------------------------------------------------------------------------
 * 段 1｜安全预置（边界 B6）：质心先落到 0，后续任何异常路径都要再覆盖它
 *      Safe preset: the centroid starts at zero, every abnormal path overwrites it
 *-----------------------------------------------------------------------------*)
FC_DL_PolygonArea := 0.0;
fCentroidX        := 0.0;
fCentroidY        := 0.0;
bCcw              := FALSE;
bDegenerate       := FALSE;
uErrorId          := 16#0000_0000;
fArea2            := 0.0;
fCxAcc            := 0.0;
fCyAcc            := 0.0;
nGuard            := 0;

(*------------------------------------------------------------------------------
 * 段 2｜点数校验（边界 B1）：上限向下钳位（多点比少点安全），下限直接拒绝
 *      Count check: clamp the upper bound down (more points is safer), reject the lower
 *-----------------------------------------------------------------------------*)
nCnt := nCount;

IF nCnt > DL_PGA_PTS_MAX THEN
    nCnt      := DL_PGA_PTS_MAX;
    uErrorId  := 16#0001_0001;
END_IF

IF nCnt < DL_PGA_PTS_MIN THEN
    (* 边界 B6：退化时给顶点算术平均，绝不返回 (0,0) *)
    (* Degenerate: return the vertex mean, never the origin *)
    IF nCnt < 1 THEN
        fCentroidX := 0.0;
        fCentroidY := 0.0;
    ELSE
        fMeanX := 0.0;
        fMeanY := 0.0;
        FOR nI := 0 TO (nCnt - 1) DO
            fMeanX := fMeanX + afX[nI];
            fMeanY := fMeanY + afY[nI];
        END_FOR
        fCentroidX := fMeanX / INT_TO_LREAL(nCnt);
        fCentroidY := fMeanY / INT_TO_LREAL(nCnt);
    END_IF
    bDegenerate := TRUE;
    uErrorId    := 16#0002_000C;
    RETURN;
END_IF

(*------------------------------------------------------------------------------
 * 段 3｜单遍累加（鞋带公式）：边权与质心权重共用同一个叉积项，只算一次
 *      Single-pass shoelace: the edge weight and the centroid weight share one cross term
 *      nJ 用 MOD nCount 闭合，nCnt >= 3 已保证除数非零，索引永不等于 nCnt
 *-----------------------------------------------------------------------------*)
FOR nI := 0 TO (nCnt - 1) DO

    nJ     := (nI + 1) MOD nCnt;
    fCross := (afX[nI] * afY[nJ]) - (afX[nJ] * afY[nI]);

    fArea2 := fArea2 + fCross;
    fCxAcc := fCxAcc + ((afX[nI] + afX[nJ]) * fCross);
    fCyAcc := fCyAcc + ((afY[nI] + afY[nJ]) * fCross);

    nGuard := nGuard + 1;

END_FOR

IF nGuard > (nCnt + 1) THEN
    (* 理论上不可达（FOR 定长），纯防御：循环计数异常即报表 *)
    (* Unreachable in theory: a bounded FOR loop cannot overrun, defence only *)
    uErrorId := 16#0001_0004;
END_IF

(*------------------------------------------------------------------------------
 * 段 4｜退化判定（边界 B3/B6）：共线或重合时面积为零，质心回退算术平均
 *      Degenerate test: zero area falls back to the vertex mean
 *-----------------------------------------------------------------------------*)
IF ABS(fArea2) <= DL_PGA_EPS THEN

    fMeanX := 0.0;
    fMeanY := 0.0;
    FOR nI := 0 TO (nCnt - 1) DO
        fMeanX := fMeanX + afX[nI];
        fMeanY := fMeanY + afY[nI];
    END_FOR

    fCentroidX  := fMeanX / INT_TO_LREAL(nCnt);
    fCentroidY  := fMeanY / INT_TO_LREAL(nCnt);
    bCcw        := FALSE;
    bDegenerate := TRUE;
    uErrorId    := 16#0002_000C;
    FC_DL_PolygonArea := 0.0;
    RETURN;

END_IF

(*------------------------------------------------------------------------------
 * 段 5｜正常路径：面积 = |fArea2| / 2，质心 = 累加 / (3 × fArea2)
 *      Normal path: area = |fArea2| / 2, centroid = accumulator / (3 × fArea2)
 *      分母用 3×fArea2 而不是 6×(fArea2/2)，少一次除法，少一次舍入
 *      bCcw 由 fArea2 的符号直接给出，不做"面积恒正后再判断"的二次推导
 *-----------------------------------------------------------------------------*)
bCcw := (fArea2 > 0.0);

fDen := DL_PGA_THREE * fArea2;

IF ABS(fDen) > DL_PGA_EPS THEN
    fCentroidX := fCxAcc / fDen;
    fCentroidY := fCyAcc / fDen;
ELSE
    (* 二次防御：段 4 已排除近零面积，此处仅防数值极端情形下的除零 *)
    (* Second defence: near-zero area was excluded in stage 4, this guards extremes *)
    fCentroidX  := 0.0;
    fCentroidY  := 0.0;
    bDegenerate := TRUE;
    uErrorId    := 16#0002_000C;
END_IF

FC_DL_PolygonArea := ABS(fArea2) / DL_PGA_TWO;
END_FUNCTION

(* ---- FC_DL_PowerFactorCalc.st ---- *)
// FC_DL_PowerFactorCalc v1.0.0
// 开源溯源：self-cleanroom / 公开公式（功率因数 = 有功/视在）
(*
  道莅工业代码库 | DL_MathData | FC_DL_PowerFactorCalc
  版本: 1.0.0 | 日期: 2026-11-23 | 轮次: R75
  功能: 功率因数计算 pf = P/S（有功/视在比），分母防零 + 领前/滞后判别；
        |pf| > 1 判测量矛盾拒收（物理不可能，疑 CT/PT 接线错误）
  邻件关系: 电能质量族 ThdCalc / HarmonicSpectrumBin（谐波畸变与频谱）——
            差异点：本件为基波功率三角比（cos φ 语义），与谐波族互不重叠
*)
FUNCTION FC_DL_PowerFactorCalc : REAL
VAR_INPUT
    fActiveKW   : REAL := 0.0;   // 有功功率 P [kW]，正=滞后感性 / Active power P [kW], positive = lagging
    fApparentKVA: REAL := 0.0;   // 视在功率 S [kVA]，域 > 0 / Apparent power S [kVA], domain > 0
    fEps        : REAL := 1.0E-6;// 判零容差 [kVA] / Zero tolerance [kVA]
END_VAR
VAR_OUTPUT
    bValid    : BOOL;            // 结果有效回执 [-] / Result validity receipt
    bLeading  : BOOL;            // 领前标志（有功为负即容性领前）[-] / Leading flag (negative P)
    uErrorId  : UDINT;           // 事件码，0 = 无事件；16#0002_1E01 = 视在为零；16#0002_1E02 = |pf|>1 矛盾 / Event code
END_VAR

// —— 段 0：全路径缺省 —— //
bValid   := FALSE;               // 有效回执预清 / Validity preset
bLeading := FALSE;               // 领前标志预清 / Leading preset
uErrorId := 16#0000;             // 事件码预清 / Event code preset
FC_DL_PowerFactorCalc := 0.0;    // 返回值缺省零 / Return default zero

// —— 段 1：非有限闸 —— //
IF (fActiveKW <> fActiveKW) OR (fApparentKVA <> fApparentKVA)
   OR (ABS(fActiveKW) >= 3.0E38) OR (ABS(fApparentKVA) >= 3.0E38) THEN
    uErrorId := 16#0002_1E01;    // 输入非有限：拒收（与视在为零共用域闸码段）/ Non-finite input: reject
    RETURN;
END_IF

// —— 段 2：分母防零闸（R4：除法前判分母） —— //
IF ABS(fApparentKVA) < fEps THEN // 视在功率近零：无法求比 / Apparent near zero: ratio undefined
    uErrorId := 16#0002_1E01;    // 信息级：分母为零 / Info level: zero denominator
    RETURN;                      // 返回零，不除 / Return zero without division
END_IF

// —— 段 3：主计算与物理矛盾闸 —— //
FC_DL_PowerFactorCalc := fActiveKW / fApparentKVA;   // pf = P/S（分母已过闸）/ pf = P/S, denominator gated
bLeading := (fActiveKW < 0.0);   // 有功为负：容性领前 / Negative P: capacitive leading
IF ABS(FC_DL_PowerFactorCalc) > 1.0 + fEps THEN      // |pf| > 1：测量矛盾 / |pf| > 1: measurement contradiction
    uErrorId := 16#0002_1E02;    // 信息级：功率三角矛盾（疑接线错误）/ Info level: power triangle contradiction
    FC_DL_PowerFactorCalc := 0.0;                    // 矛盾值不外发，返回零 / Contradictory value suppressed
    RETURN;
END_IF
bValid := TRUE;                  // 有效回执 / Validity receipt
END_FUNCTION

(* ---- FC_DL_PowIntSat.st ---- *)
(*
    FC_DL_PowIntSat —— 整数幂 Safe 族防御包装（指数钳位 [0,63] + 显式符号分支 + 溢出饱和）
    ------------------------------------------------------------------
    分类      : DL_MathData / Math-Power
    前缀      : FC_DL_
    版本      : 1.0.1
    来源标签  : iec-std-wrapper（T0）
    溯源      : IEC 61131-3 标准语义的道莅防御性实现
                （纯循环乘法实现，不依赖 EXPT 浮点路径，无幂运算符；
                  未复制任何闭源厂商源码）
    平台      : 纯 IEC 61131-3，CODESYS / TwinCAT / InoProShop 通用
    分工声明  : 与存量 FC_DL_ExptEx / FC_DL_FactorialSat 分工——ExptEx 为浮点
                任意底任意指数码位族（委托 EXPT），本件为整数指数幂的 Safe 族
                口径（循环乘 + 预检饱和）；FactorialSat 只做阶乘口径。
    作者      : 道莅代码库 · PLC 编程专家（R57）
    ------------------------------------------------------------------
    功能说明  : 求 fBase 的 nExp 整数次幂。四段式防御（R45）：底数/指数非有限
                双判据拦截；nExp 钳位 [0, 63]（极限值→可表性反算，R63：2^63
                约 9.22E18，最大底数 1.79E308 时 2 次幂即越界，由乘法预检饱和
                兜底，63 为指数域钳位上界）；底 0 且 0 次幂判错误（返回 0）；
                负底符号按奇偶显式分支（|底| 循环乘，符号末段乘回）；每次乘法
                前做 acc > MAX/|底| 预检防 Inf，超界饱和。
    错误码    : 0000 正常 / 16#0002_0001 入参非有限已归零 / 16#0002_0002 指数已钳位 / 16#0002_0003 底 0 的 0 次幂 / 16#0002_0006 结果已饱和
    修订记录  : 2026-11-21 v1.0.0 首次入库（R57 批 2 · 序号 10）
                2026-11-21 v1.0.1 R58 返修：段 4 饱和置码 0206 原为无条件，会
                覆盖先发事件 0202（指数钳位）；补首事件闸对齐段 5 口径；95~97
                行 bError/bValid/bClamped 保持无条件（标志级聚合，码级唯一）。
*)
FUNCTION FC_DL_PowIntSat : LREAL
VAR_INPUT
    fBase : LREAL; // 底数实数 [无量纲] / the base real value [dimensionless]
    nExp  : INT;   // 整数指数 [次]，钳位 [0, 63] / the integer exponent, clamped to zero through sixty three
END_VAR
VAR_OUTPUT
    eErr     : UDINT; // 错误码，0 = 正常 / error code, zero is ok
    bError   : BOOL;  // 出错标志，eErr 非 0 时为真 / error flag, true when eErr is nonzero
    bValid   : BOOL;  // 结果是否为真实值，钳位/饱和降级时为假 / the result is the true value, false when degraded
    bClamped : BOOL;  // 本次调用发生指数或幅值钳位 [-] / an exponent or magnitude clamp happened this call
END_VAR
VAR
    lrMag  : LREAL; // 幅值累乘量 [无量纲] / the magnitude accumulator [dimensionless]
    lrAbB  : LREAL; // 底数绝对值 [无量纲] / the base magnitude [dimensionless]
    nI     : INT;   // 循环计数 [次] / the loop counter
    bNeg   : BOOL;  // 结果应为负（负底奇次幂）[-] / the result should be negative, an odd power of a negative base
END_VAR
VAR CONSTANT
    DL_POW_EXPMAX : INT   := 63;                  // 指数钳位上界 [次]（R63）/ the exponent clamp bound
    DL_POW_MAGMAX : LREAL := 1.7976931348623157E308; // LREAL 可表上界 [无量纲] / the representable magnitude bound
END_VAR

// 段 1｜返回值与错误状态预置安全值（四段式第一段，R45）/ segment 1, preset the return and error states
FC_DL_PowIntSat := 0.0; // 返回值预置安全值 0.0 / preset the return to the safe zero
eErr     := 16#0000_0000; // 错误码预置正常 / preset the code to ok
bError   := FALSE; // 错误标志预置假 / preset the error flag false
bValid   := TRUE; // 有效标志预置真 / preset the valid flag true
bClamped := FALSE; // 钳位标志预置假 / preset the clamp flag false

// 段 2｜非有限拦截（双判据）：命中直接早退 / segment 2, the non finite interception
IF (fBase <> fBase) OR ((fBase - fBase) <> (fBase - fBase)) THEN // 底数非有限 / a non finite base
    eErr   := 16#0002_0001; // 信息级：底数非有限已归零 / informational, a non finite base zeroed
    bError := TRUE; // 置错误标志 / raise the error flag
    bValid := FALSE; // 输出不可用 / the output void
    RETURN; // 返回预置安全值 0.0 / return the preset safe zero
END_IF

// 段 3｜指数钳位与底 0 的 0 次幂判定 / segment 3, the exponent clamp and the zero base zero power
IF nExp < 0 THEN // 负指数越下界 / a negative exponent
    nExp     := 0; // 钳到 0 / clamp to zero
    eErr     := 16#0002_0002; // 信息级：指数已钳位 / informational, the exponent clamped
    bError   := TRUE; // 置错误标志 / raise the error flag
    bValid   := FALSE; // 钳位结果非真实值 / the clamped result is not the true value
    bClamped := TRUE; // 置钳位标志 / raise the clamp flag
ELSIF nExp > DL_POW_EXPMAX THEN // 越上界 / above the bound
    nExp     := DL_POW_EXPMAX; // 钳到上界 / clamp to the bound
    eErr     := 16#0002_0002; // 信息级：指数已钳位 / informational, the exponent clamped
    bError   := TRUE; // 置错误标志 / raise the error flag
    bValid   := FALSE; // 钳位结果非真实值 / the clamped result is not the true value
    bClamped := TRUE; // 置钳位标志 / raise the clamp flag
END_IF
IF (fBase = 0.0) AND (nExp = 0) THEN // 底 0 的 0 次幂（数学未定义，判错误）/ the zero base zero power, undefined
    eErr   := 16#0002_0003; // 错误级：底 0 的 0 次幂返回 0 / error grade, the zero base zero power returns zero
    bError := TRUE; // 置错误标志 / raise the error flag
    bValid := FALSE; // 输出不可用 / the output void
    RETURN; // 返回预置安全值 0.0 / return the preset safe zero
END_IF
IF fBase = 0.0 THEN // 底 0 的正整数幂恒为 0 / a zero base with a positive power is zero
    RETURN; // 返回安全值 0.0，标志保持正常 / return the safe zero, the flags stay ok
END_IF

// 段 4｜幅值循环乘 + 预检饱和 + 负底奇偶符号显式分支 / segment 4, the magnitude loop with the pre-check saturation and the explicit sign branch
lrAbB := ABS(fBase); // 底数绝对值 / the base magnitude
bNeg  := (fBase < 0.0) AND ((nExp MOD 2) = 1); // 负底且奇次幂为负（nExp 非负，MOD 合法）/ negative when an odd power of a negative base
lrMag := 1.0; // 幅值从 1 起乘 / the magnitude starts at one
FOR nI := 1 TO nExp DO // 逐次乘（nExp 已钳 ≤63，循环有界）/ the bounded loop
    IF lrMag > DL_POW_MAGMAX / lrAbB THEN // 乘前预检防 Inf（除子为正底绝对值已证大于零）/ the pre-check against infinity
        lrMag    := DL_POW_MAGMAX; // 幅值饱和到可表上界 / saturate the magnitude
        IF eErr = 16#0000_0000 THEN // 首事件优先置码（对齐段 5 闸式，v1.0.1）/ the first event keeps the code, aligned with segment five
            eErr     := 16#0002_0006; // 信息级：结果已饱和 / informational, the result saturated
        END_IF
        bError   := TRUE; // 置错误标志（标志级无条件聚合）/ raise the error flag unconditionally
        bValid   := FALSE; // 饱和结果非真实值 / the saturated result is not the true value
        bClamped := TRUE; // 置钳位标志 / raise the clamp flag
        EXIT; // 提前出循环 / leave the loop early
    END_IF
    lrMag := lrMag * lrAbB; // 幅值累乘 / accumulate the magnitude
END_FOR
IF bNeg THEN // 负底奇次幂符号乘回（显式分支，边界十）/ the sign multiplied back, the explicit branch
    FC_DL_PowIntSat := -lrMag; // 负结果 / the negative result
ELSE // 正结果（含负底偶次幂）/ the positive result, including an even power of a negative base
    FC_DL_PowIntSat := lrMag; // 正结果 / the positive result
END_IF

// 段 5｜结果非有限复核兜底（防御纵深，正常路径不可达）/ segment 5, the result recheck as defense in depth
IF (FC_DL_PowIntSat <> FC_DL_PowIntSat) OR ((FC_DL_PowIntSat - FC_DL_PowIntSat) <> (FC_DL_PowIntSat - FC_DL_PowIntSat)) THEN // 结果非有限 / a non finite result
    FC_DL_PowIntSat := 0.0; // 兜底安全值 / the bottom-line safe value
    IF eErr = 16#0000_0000 THEN // 首事件优先置码 / the first event keeps the code
        eErr   := 16#0002_0001; // 信息级：结果非有限已归零 / informational, a non finite result zeroed
        bError := TRUE; // 置错误标志 / raise the error flag
        bValid := FALSE; // 输出不可用 / the output void
    END_IF
END_IF
END_FUNCTION

(* ---- FC_DL_PwrDbToRatio.st ---- *)
(*
    FC_DL_PwrDbToRatio —— 功率型分贝到线性功率比换算
    ------------------------------------------------------------------
    分类      : DL_MathData / Log
    前缀      : FC_DL_
    版本      : 1.0.0
    溯源      : IEC 61131-3 标准语义的道莅防御性实现
                （接口语义由 IEC 61131-3 定义，内部委托平台内建 EXPT，
                  外围统一错误码 / 钳位 / 双语文档；clean-room 重写，
                  未复制任何闭源厂商源码，参考实现仅限 MIT/Apache 许可）
    平台      : 纯 IEC 61131-3，CODESYS / TwinCAT / InoProShop 通用
    作者      : 道莅代码库 · PLC编程专家（R17）
    ------------------------------------------------------------------
    功能说明  : 功率型分贝转过线性功率比，按 P = 10^(dB/10) 实现，指数运算委托平台内建 EXPT，
                10 为功率型换算因子（与幅值型 20 严格区分，禁混用），不重实现指数内核；
                非有限输入判为故障级 16#0001_02D6，返回 1.0（功率比中性值）；
                |dB| 超 380.0 dB 硬限时按方向饱和至 1.0E38 / 1.0E-38，置信息级 16#0001_01F0；
                硬限取 380.0 dB 而非 400.0 dB 的理由：功率型 400 dB 对应比值 10^40，
                超出 REAL 最大有限值 3.402823E38，饱和值本身不可表；380 dB 对应 10^±38，两端均可表；
                钳位方向：双侧饱和（dB 域 ±380.0 dB，比值域 1.0E-38 ~ 1.0E38）。
    错误码    : 16#0001_01F0 dB 值超 ±380.0 dB 硬限，已按方向饱和——信息级，正常防御
                16#0001_01F1 预留禁用（信息级，不得挪用）
                16#0001_02D6 非有限输入（NaN 或 ±INF）——故障级，返回 1.0
                16#0001_02D7 预留禁用（故障级，不得挪用）
                16#0001_02D8 预留禁用（故障级，不得挪用）
    状态机    : R6 标注 N/A —— 本组件为纯函数无顺序状态机，无 CASE 可写，非法状态不可能出现，故以本节说明替代 ELSE 兜底
    修订记录  : 2026-11-16 v1.0.0 首次入库（R17）
*)
FUNCTION FC_DL_PwrDbToRatio : REAL
VAR_INPUT
    fDb : REAL; // 功率型分贝值，建议域 −380.0~+380.0 [dB] / power decibel value, suggested domain -380.0..+380.0 [dB]
END_VAR
VAR_OUTPUT
    eErr   : UDINT; // 错误码，0=正常 / error id, 0=ok
    bError : BOOL;  // 是否出错，eErr 非 0 时为 TRUE / error flag, TRUE when eErr is nonzero
    bValid : BOOL;  // 输出是否有效可用 / output valid flag
END_VAR
VAR CONSTANT
    DL_DB_PWR_DIV     : REAL := 10.0;     // 功率型 dB 换算除子（10·log10 的逆向） [dB] / power dB divisor, inverse of 10*log10 [dB]
    DL_DB_TEN         : REAL := 10.0;     // 幂运算底数 10 [无量纲] / power base 10 [dimensionless]
    DL_DB_PWR_LIMIT   : REAL := 380.0;    // 功率型 dB 域双侧硬限，对应比值 10^±38（400 dB 会超出 REAL 域） [dB] / power dB hard limit, ratio 10^+/-38 [dB]
    DL_RATIO_NEUTRAL  : REAL := 1.0;      // 功率比中性值（0 dB 对应值，故障缺省返回） [比] / neutral power ratio (0 dB), fault default [ratio]
    DL_PWR_RATIO_MAX  : REAL := 1.0E38;   // 功率比上限 10^38，REAL 域可表 [比] / power ratio upper bound 10^38 [ratio]
    DL_PWR_RATIO_MIN  : REAL := 1.0E-38;  // 功率比下限 10^-38，REAL 域可表 [比] / power ratio lower bound 10^-38 [ratio]
    DL_REAL_INF_GUARD : LREAL := 4.0E38;  // REAL 域 ±INF 判定阈值，高于 REAL 最大有限值 3.402823E38 [无量纲] / REAL +/-INF guard above max finite REAL
END_VAR
VAR
    bNonFinite : BOOL; // 非有限（NaN 或 ±INF）判定结果 / non-finite (NaN or +/-INF) detection result
END_VAR

// 段 1｜返回值与错误状态预置 / segment 1, preset return value and error status
FC_DL_PwrDbToRatio := DL_RATIO_NEUTRAL; // 故障缺省返回 1.0 功率比中性值 [比] / fault default 1.0 neutral power ratio [ratio]
eErr   := 0;     // 预置无错误 / preset no error
bError := FALSE; // 预置无故障 / preset no fault
bValid := FALSE; // 预置输出无效，通过非有限闸后置位 / preset invalid, set TRUE after the non-finite gate

// 段 2｜非有限防御闸 / segment 2, non-finite guard
bNonFinite := (fDb <> fDb) OR (fDb > DL_REAL_INF_GUARD) OR (fDb < -DL_REAL_INF_GUARD); // 非有限判定（NaN 自不等 + 安全幅值判 ±INF） [dB] / non-finite check (NaN by self-inequality, +/-INF by safe magnitude) [dB]
IF bNonFinite THEN
    eErr := 16#0001_02D6; // 非有限输入故障码 / non-finite input fault id
    bError := TRUE;       // 置故障标志 / raise error flag
    bValid := FALSE;      // 输出不可用 / output not usable
    RETURN;               // 故障级提前返回，保持缺省 1.0 / early return on fault, keep default 1.0
END_IF

// 段 3｜dB 域硬限双侧饱和 / segment 3, two-sided dB domain saturation
IF fDb > DL_DB_PWR_LIMIT THEN
    FC_DL_PwrDbToRatio := DL_PWR_RATIO_MAX; // 正超饱和至功率比上限 1.0E38 [比] / positive overflow saturates to power ratio upper bound 1.0E38 [ratio]
    eErr := 16#0001_01F0;                   // 信息级：dB 超限已饱和，正常防御 / info level: dB exceeded the limit and saturated, normal defence
    bError := FALSE;                        // 信息级不置故障 / info level never raises fault
    bValid := TRUE;                         // 饱和值本身有效可用 / the saturated value itself is valid
    RETURN;                                 // 饱和即出口，不进入幂运算 / saturation is the exit, no power computation
END_IF
IF fDb < -DL_DB_PWR_LIMIT THEN
    FC_DL_PwrDbToRatio := DL_PWR_RATIO_MIN; // 负超饱和至功率比下限 1.0E-38 [比] / negative overflow saturates to power ratio lower bound 1.0E-38 [ratio]
    eErr := 16#0001_01F0;                   // 同一业务语义复用同一信息码 / same business semantics reuses the same info id
    bError := FALSE;                        // 信息级不置故障 / info level never raises fault
    bValid := TRUE;                         // 饱和值本身有效可用 / the saturated value itself is valid
    RETURN;                                 // 饱和即出口，不进入幂运算 / saturation is the exit, no power computation
END_IF

// 段 4｜主体幂运算与结果复检（末段） / segment 4, main power computation and result re-check (final)
FC_DL_PwrDbToRatio := EXPT(DL_DB_TEN, fDb / DL_DB_PWR_DIV); // 域内委托内建 EXPT 计算 10^(dB/10) [比] / in-domain delegate to built-in EXPT for 10^(dB/10) [ratio]
IF (FC_DL_PwrDbToRatio <> FC_DL_PwrDbToRatio) OR (FC_DL_PwrDbToRatio > DL_PWR_RATIO_MAX) OR (FC_DL_PwrDbToRatio < DL_PWR_RATIO_MIN) THEN // 结果复检：NaN 自不等 + 双侧越界（±INF 亦被幅值界捕获） [比] / result re-check: NaN by self-inequality plus two-sided overflow, +/-INF also caught by the magnitude bounds [ratio]
    IF fDb >= 0.0 THEN
        FC_DL_PwrDbToRatio := DL_PWR_RATIO_MAX; // 按输入符号方向饱和至上限 [比] / saturate upward following the input sign [ratio]
    ELSE
        FC_DL_PwrDbToRatio := DL_PWR_RATIO_MIN; // 按输入符号方向饱和至下限 [比] / saturate downward following the input sign [ratio]
    END_IF
    eErr := 16#0001_01F0; // 溢出行为差异复用同一信息码，不另立码 / platform overflow difference reuses the same info id, no extra code
    bError := FALSE;      // 信息级不置故障 / info level never raises fault
    bValid := TRUE;       // 饱和值本身有效可用 / the saturated value itself is valid
    RETURN;               // 复检出口 / exit after the re-check
END_IF
eErr   := 0;     // 域内无错误 / in-domain, no error
bError := FALSE; // 信息级不置故障 / info level never raises fault
bValid := TRUE;  // 域内输出有效可用 / in-domain output is valid
END_FUNCTION

(* ---- FC_DL_QuadPolyFit.st ---- *)
(*
  ==================================================================
  组件名 Component  : FC_DL_QuadPolyFit
  分类   Category   : DL_MathData
  版本   Version    : 1.0.1
  功能   Purpose    : 二次多项式最小二乘拟合 y = a0 + a1*x + a2*x²：构造 3×3
                      正规方程（Σ 0~4 阶矩 + 0~2 阶矩与 y 的混合矩），列主元
                      Gauss 消元求解。主元 |p| < 1E-10 判奇异：不输出系数、
                      bValid=FALSE、码 03（不静默给退化系数）。三重 FOR 均
                      以常量封顶（消元 2 轮 × 选行 3 行 × 回代 3 元）。
  来源   Source     : t2-1-lgf-math（数学族：正规方程 + 列主元消元为公开
                      数值方法口径，实现零源码复制）
  互引   Cross-ref  : FC_DL_LinearRegression2Var（同族低阶拟合原子，本件为其
                      二次扩展，共用「矩累加 + 正规方程」方法论）
  平台   Platform   : 纯 IEC 61131-3 四则 + ABS/TRUNC，三平台通用
  依赖   Depends    : 无 DL_ 内部依赖；无标准库
  设计偏差 Deviation: nCount > 数组实际长度时按长度钳位接管（同族口径，头注
                      声明，不静默越界，见码位反证）；y = a0+a1x+a2x² 系数
                      排序为「常数项在前」，返回值 = fA0（名实双出口）。
  红线   Redline    : R1 零全局/VAR_EXTERNAL/R2 零 %I/%Q/R3 纯 IEC 标准
                      R4 点数闸 + 元素级非有限闸 + 矩溢出非有限复核 +
                      主元闸（禁除以近零）/R5 全变量双语同行注释
                      R6 纯函数无状态机（CASE 不适用）/R7 无定时器与沿检测
                      R8 阈值与循环界全常量化
  错误码 Codes      : 01【失效级】点数不足（钳位后 nCount < 3），返回 0
                      02【失效级】任一 x/y 非有限或矩累加溢出为非有限
                      03【失效级】正规方程奇异（列主元 < 1E-10），不输出系数
  码位反证 Note     : 01/02/03 分立依据（R90）：01 在计数面、02 在数据面、
                      03 在数值结构面可观测；03 若并入 02，则「给不给退化
                      系数」这一行为差异将不可观测，故必须分立。
  验收   Acceptance : V1 完美 y=x² 采样 → a2≈1，a0/a1≈0 ｜ V2 2 点 → 码 01
                      ｜ V3 含 NaN → 码 02 ｜ V4 全部 x 相同（奇异）→ 码 03
                      ｜ V4b 仅两个相异 x（秩 2，舒尔补奇异）→ 码 03（v1.0.1）
                      ｜ V5 带噪数据 → 残差递减于线性拟合
  变更   Revision   : 2026-11-22  v1.0.0  R66 首版（编码阶段批 2 序 6）
                      2026-11-22  v1.0.1  R67 点修（M2+L1）：段 7 回代前补
                      舒尔补主元闸 aM[2,2]（两相异 x 值正规方程秩 2 场景，
                      除零 NaN/Inf 原错归码 02 → 提前归码 03）；段 4 ABS 溢
                      出复核由 s4/t2 扩展至 s1/s2/s3/t0/t1 全部矩量。
  ==================================================================
*)
FUNCTION FC_DL_QuadPolyFit : LREAL
VAR_INPUT
    aX     : ARRAY[*] OF LREAL;  // 自变量数组 [物理单位] / the abscissa array
    aY     : ARRAY[*] OF LREAL;  // 因变量数组 [物理单位] / the ordinate array
    nCount : UDINT;              // 参与拟合点数 [个]，超出数组长度按长度钳位 / the sample count, clamped to the array length
END_VAR
VAR_OUTPUT
    fA0    : LREAL;  // 拟合系数常数项 [物理单位]（y = a0 + a1*x + a2*x²）/ the constant coefficient
    fA1    : LREAL;  // 拟合系数一次项 [斜率] / the linear coefficient
    fA2    : LREAL;  // 拟合系数二次项 [1/斜率单位] / the quadratic coefficient
    bValid : BOOL;   // 系数可用标志 [-] / the coefficients usable flag
    nErrId : UDINT;  // 错误码，0=正常，01/02/03 见头注 [码] / the error code [code]
END_VAR
VAR
    s0     : LREAL;  // Σx^0 矩 [个] / the zeroth moment
    s1     : LREAL;  // Σx^1 矩 / the first moment
    s2     : LREAL;  // Σx^2 矩 / the second moment
    s3     : LREAL;  // Σx^3 矩 / the third moment
    s4     : LREAL;  // Σx^4 矩 / the fourth moment
    t0     : LREAL;  // Σy 矩 [物理单位] / the y moment
    t1     : LREAL;  // Σxy 矩 / the xy moment
    t2     : LREAL;  // Σx²y 矩 / the x squared y moment
    fx     : LREAL;  // 当前 x 工作寄存器 / the current x working register
    fy     : LREAL;  // 当前 y 工作寄存器 / the current y working register
    fx2    : LREAL;  // 当前 x² 工作寄存器 / the current x squared register
    aM     : ARRAY[0..2, 0..2] OF LREAL; // 正规方程系数矩阵 / the normal equation coefficient matrix
    aR     : ARRAY[0..2] OF LREAL;       // 正规方程右端向量 / the normal equation right hand vector
    aSol   : ARRAY[0..2] OF LREAL;       // 解向量工作寄存器 / the solution working vector
    uUsed  : UDINT;  // 钳位后实际点数 [个] / the used count after clamping
    uLenX  : UDINT;  // aX 实际长度 [个] / the actual length of aX
    uLenY  : UDINT;  // aY 实际长度 [个] / the actual length of aY
    uLen   : UDINT;  // 双数组共同安全长度 [个] / the common safe length
    i      : UDINT;  // 采样累加循环变量 / the accumulation loop index
    k      : DINT;   // 消元主轮变量，0~1 / the elimination pass index
    p      : DINT;   // 选主元行扫描变量 / the pivot row scan index
    r      : DINT;   // 消元行扫描变量 / the elimination row scan index
    c      : DINT;   // 消元列扫描变量 / the elimination column scan index
    fPivot : LREAL;  // 当轮主元值 / the current pivot value
    iMax   : DINT;   // 当轮主元所在行 / the pivot row of this pass
    fFac   : LREAL;  // 消元因子 / the elimination factor
    fTmp   : LREAL;  // 行交换临时量 / the row swap temporary
END_VAR
VAR CONSTANT
    QPF_PIV_MIN   : LREAL := 1.0E-10;             // 主元奇异阈值 [无量纲] / the singular pivot threshold
    QPF_PTS_MIN   : UDINT := UDINT#3;             // 二次拟合最少点数 [个] / the minimum points for a quadratic fit
    QPF_FIN_MAX   : LREAL := 1.7976931348623157E308; // LREAL 有限上限 / the finite LREAL limit
    QPF_ELIM_PASS : DINT := 2;                    // 消元主轮数（3×3 方程组）/ the elimination passes for a 3 by 3 system
    QPF_DIM       : DINT := 3;                    // 方程组维数 / the system dimension
    QPF_ERR_NONE  : UDINT := 16#0000_0000;        // 无错误 [码] / no error [code]
    QPF_ERR_PTS   : UDINT := 16#0000_0001;        // 码 01：点数不足 / code 01, too few points
    QPF_ERR_NAN   : UDINT := 16#0000_0002;        // 码 02：非有限 / code 02, non finite
    QPF_ERR_SING  : UDINT := 16#0000_0003;        // 码 03：奇异 / code 03, singular
END_VAR

// 段 1｜输出预置 / segment 1, preset the outputs
FC_DL_QuadPolyFit := 0.0;  // 失效缺省返回 0（=fA0 缺省）/ fault default returns zero
fA0    := 0.0;             // 系数预置 0（奇异不输出退化系数，头注口径）/ preset zero, no degenerate coefficients on singularity
fA1    := 0.0;
fA2    := 0.0;
bValid := FALSE;           // 预置不可用 / preset unusable
nErrId := QPF_ERR_NONE;    // 预置无错误 / preset no error
s0 := 0.0; s1 := 0.0; s2 := 0.0; s3 := 0.0; s4 := 0.0;  // 矩累加器清零 / clear the moment accumulators
t0 := 0.0; t1 := 0.0; t2 := 0.0;                        // 混合矩累加器清零 / clear the mixed moment accumulators

// 段 2｜数组长度闸与点数闸（结构 RETURN 早退）/ segment 2, the length and count gates
IF UPPER_BOUND(aX, 1) >= 0 THEN                          // 防御性变长上界检查 / defensive bound check
    uLenX := DINT_TO_UDINT(1 + UPPER_BOUND(aX, 1) - LOWER_BOUND(aX, 1));  // aX 长度 / the aX length
ELSE
    uLenX := UDINT#0;
END_IF
IF UPPER_BOUND(aY, 1) >= 0 THEN
    uLenY := DINT_TO_UDINT(1 + UPPER_BOUND(aY, 1) - LOWER_BOUND(aY, 1));  // aY 长度 / the aY length
ELSE
    uLenY := UDINT#0;
END_IF
IF uLenX < uLenY THEN                                    // 双数组取共同安全长度 / the common safe length
    uLen := uLenX;
ELSE
    uLen := uLenY;
END_IF
uUsed := nCount;                                         // 先取原始点数 / take the raw count
IF uUsed > uLen THEN
    uUsed := uLen;                                       // 超长钳位接管（头注偏差声明）/ clamp, documented deviation
END_IF
IF uUsed < QPF_PTS_MIN THEN                              // 点数不足（码 01）/ too few points, code 01
    nErrId := QPF_ERR_PTS;
    RETURN;
END_IF

// 段 3｜矩累加：元素级非有限闸（码 02）+ 下标闸已证（uUsed ≤ uLen）
//      segment 3, the moment accumulation with the per element finite gate
FOR i := 0 TO UDINT_TO_DINT(uUsed) - 1 DO                // 有界 FOR / the bounded loop
    fx := aX[i];                                         // 当前 x / the current x
    fy := aY[i];                                         // 当前 y / the current y
    IF (fx <> fx) OR (fy <> fy) OR (ABS(fx) > QPF_FIN_MAX) OR (ABS(fy) > QPF_FIN_MAX) THEN
        nErrId := QPF_ERR_NAN;                           // 码 02：非有限元素 / code 02, non finite element
        RETURN;                                          // 结构早退 / structural early return
    END_IF
    fx2 := fx * fx;                                      // 当前 x² / the current x squared
    s0 := s0 + 1.0;                                      // 零阶矩累加 / the zeroth moment
    s1 := s1 + fx;                                       // 一阶矩 / the first moment
    s2 := s2 + fx2;                                      // 二阶矩 / the second moment
    s3 := s3 + fx2 * fx;                                 // 三阶矩 / the third moment
    s4 := s4 + fx2 * fx2;                                // 四阶矩 / the fourth moment
    t0 := t0 + fy;                                       // Σy / the y moment
    t1 := t1 + fx * fy;                                  // Σxy / the xy moment
    t2 := t2 + fx2 * fy;                                 // Σx²y / the x squared y moment
END_FOR

// 段 4｜矩溢出非有限复核（码 02）：极端量级下累加可能溢出 Inf，先闸后入阵
//      segment 4, the overflow recheck on the moments before entering the matrix
IF (s0 <> s0) OR (s1 <> s1) OR (s2 <> s2) OR (s3 <> s3) OR (s4 <> s4)
   OR (t0 <> t0) OR (t1 <> t1) OR (t2 <> t2)
   OR (ABS(s1) > QPF_FIN_MAX) OR (ABS(s2) > QPF_FIN_MAX)     // v1.0.1 扩展 / extended in v1.0.1
   OR (ABS(s3) > QPF_FIN_MAX) OR (ABS(s4) > QPF_FIN_MAX)     // v1.0.1 扩展 / extended in v1.0.1
   OR (ABS(t0) > QPF_FIN_MAX) OR (ABS(t1) > QPF_FIN_MAX)     // v1.0.1 扩展 / extended in v1.0.1
   OR (ABS(t2) > QPF_FIN_MAX) THEN
    nErrId := QPF_ERR_NAN;
    RETURN;
END_IF

// 段 5｜构造 3×3 正规方程 / segment 5, build the 3 by 3 normal equations
aM[0,0] := s0;  aM[0,1] := s1;  aM[0,2] := s2;           // 第一行 [a0 系数] / the first row
aM[1,0] := s1;  aM[1,1] := s2;  aM[1,2] := s3;           // 第二行 [a1 系数] / the second row
aM[2,0] := s2;  aM[2,1] := s3;  aM[2,2] := s4;           // 第三行 [a2 系数] / the third row
aR[0] := t0;  aR[1] := t1;  aR[2] := t2;                 // 右端向量 / the right hand side

// 段 6｜列主元 Gauss 消元（常量封顶双重 FOR）/ segment 6, column pivoted elimination
FOR k := 0 TO QPF_ELIM_PASS - 1 DO                       // 逐主轮 / pass by pass
    fPivot := ABS(aM[k,k]);                              // 初选对角元 / seed with the diagonal
    iMax := k;                                           // 初选行 / the seeded row
    FOR p := k + 1 TO QPF_DIM - 1 DO                     // 列内选主元 / the column pivot scan
        IF ABS(aM[p,k]) > fPivot THEN
            fPivot := ABS(aM[p,k]);                      // 更大主元 / the larger pivot
            iMax := p;                                   // 主元行 / the pivot row
        END_IF
    END_FOR
    IF fPivot < QPF_PIV_MIN THEN                         // 主元闸（码 03）：禁除以近零 / the pivot gate
        nErrId := QPF_ERR_SING;
        RETURN;                                          // 不输出系数（头注口径）/ no coefficients published
    END_IF
    IF iMax <> k THEN                                    // 行交换 / the row swap
        FOR c := 0 TO QPF_DIM - 1 DO                     // 交换系数行 / swap the coefficient row
            fTmp := aM[k,c];  aM[k,c] := aM[iMax,c];  aM[iMax,c] := fTmp;
        END_FOR
        fTmp := aR[k];  aR[k] := aR[iMax];  aR[iMax] := fTmp;  // 交换右端 / swap the right hand side
    END_IF
    FOR r := k + 1 TO QPF_DIM - 1 DO                     // 消元行扫描 / the elimination row scan
        fFac := aM[r,k] / aM[k,k];                       // 除数 = 主元，已闸 ≥ 1E-10 / the divisor is the gated pivot
        FOR c := k TO QPF_DIM - 1 DO                     // 行内消元 / the in row elimination
            aM[r,c] := aM[r,c] - fFac * aM[k,c];
        END_FOR
        aR[r] := aR[r] - fFac * aR[k];                   // 右端同步消元 / eliminate the right hand side too
    END_FOR
END_FOR

// 段 7｜回代前舒尔补主元闸（v1.0.1）：消元主轮仅覆盖第 0/1 列，aM[2,2] 为舒
//      尔补未经闸——两个相异 x 值（正规方程秩 2，传感器两态卡值可达）时
//      aM[2,2]=0，回代除零出 NaN/Inf 原落段 8 码 02，与头注码 03（奇异）
//      归因错位，故回代前按码 03 提前拦截
//      segment 7, the Schur complement pivot gate before back substitution
IF ABS(aM[2,2]) < QPF_PIV_MIN THEN                        // 舒尔补主元闸（双精度口径，阈同主元闸）/ the Schur complement pivot gate
    nErrId := QPF_ERR_SING;                               // 码 03：正规方程秩 2 奇异 / code 03, rank two singular
    RETURN;                                               // 不输出系数（bValid 段 1 已预置 FALSE）/ no coefficients published
END_IF
aSol[2] := aR[2] / aM[2,2];                              // a2 回代解（舒尔补已闸）/ the quadratic unknown, Schur complement gated
aSol[1] := (aR[1] - aM[1,2] * aSol[2]) / aM[1,1];        // a1 回代解 / the linear unknown
aSol[0] := (aR[0] - aM[0,1] * aSol[1] - aM[0,2] * aSol[2]) / aM[0,0];  // a0 回代解 / the constant unknown

// 段 8｜解的非有限复核（码 02）与出口 / segment 8, the solution finiteness recheck and exit
IF (aSol[0] <> aSol[0]) OR (aSol[1] <> aSol[1]) OR (aSol[2] <> aSol[2])
   OR (ABS(aSol[2]) > QPF_FIN_MAX) THEN
    nErrId := QPF_ERR_NAN;                               // 极端病态下回代仍可能溢出 / the substitution can still overflow in extreme ill conditioning
    RETURN;
END_IF
fA0 := aSol[0];                                          // 发布常数项 / publish the constant
fA1 := aSol[1];                                          // 发布一次项 / publish the linear term
fA2 := aSol[2];                                          // 发布二次项 / publish the quadratic term
bValid := TRUE;                                          // 系数可用 / the coefficients are usable
FC_DL_QuadPolyFit := fA0;                                // 返回值 = fA0（R191 名实双出口，头注偏差声明）/ the return mirrors fA0
END_FUNCTION

(* ---- FC_DL_QuadraticSolve.st ---- *)
(*
  ==================================================================
  组件名 Component  : FC_DL_QuadraticSolve
  分类   Category   : DL_MathData
  复杂度 Complexity  : 轻
  版本   Version    : 1.0.0
  功能   Purpose    : 二次方程 a·x² + b·x + c = 0 实根求解。判别式三域分档：
                      D > eps 两实根（x1 ≥ x2）、|D| ≤ eps 重根、D < -eps 无
                      实根（nRoots = 0，非故障）；a ≈ 0 退化线性分支（b ≈ 0
                      再分恒成立/无解）；全程浮点禁等号，用 ABS 阈值。
                      OSCAT Basic 数值域公开语义 clean-room。
  来源   Source     : T1-1-oscat-basic（数值域公开语义）
  溯源   Origin     : 二次方程求根公式为公开数学语义，clean-room 自研实现，
                      未复制 OSCAT 或任何厂商私有库源码。
  平台   Platform   : 纯 IEC 61131-3，CODESYS / TwinCAT / InoProShop 通用
  分工声明 Split     : 与 FC_DL_SimpsonQuad 分工——后者做数值积分，本件做
                      二次方程解析求根。
  作者   Author     : 道莅代码库 · PLC 编程专家（R59）
  ------------------------------------------------------------------
  边界 Boundary     :
                      一 非有限入参闸（自反双判据，三参数全覆盖）：命中置
                         bError 早退，输出安全侧零（四段式 R45）；
                      二 除零闸：线性分支除 b、求根除 2a 前强制 |系数| ≥ eps
                         判据（已由分支条件保证，代码内再显式闸一层）；
                      三 SQRT 域闸：仅 D ≥ 0 才开方（判据前置）；
                      四 nRoots = -1 表示 a = b = 0 且 c = 0 恒成立（全 x 均
                         为解），nRoots = 0 无实根，均为信息级非故障；
                      五 无全局变量、无外部变量声明、无物理地址寻址。
  修订记录 Revision  :
    2026-11-21  v1.0.0  R59 首版（批 1 · 序号 5）
  ==================================================================
*)

FUNCTION FC_DL_QuadraticSolve : BOOL
VAR_INPUT
    fA : LREAL := 0.0; // 二次项系数 [无量纲] / the quadratic coefficient
    fB : LREAL := 0.0; // 一次项系数 [无量纲] / the linear coefficient
    fC : LREAL := 0.0; // 常数项 [无量纲] / the constant term
END_VAR
VAR_OUTPUT
    fX1    : LREAL := 0.0; // 实根一（两根时较大者）[无量纲] / the real root one, the larger when two roots
    fX2    : LREAL := 0.0; // 实根二 [无量纲] / the real root two
    nRoots : DINT  := 0;   // 实根个数：0 无 / 1 重根或线性 / 2 两根 / -1 恒成立 [个] / the real root count, minus one means identity
    bLinear: BOOL := FALSE; // a ≈ 0 退化线性分支受理 [-] / the degenerate linear branch accepted
    bValid : BOOL := FALSE; // 结果可用标志 [-] / the result usable flag
    bError : BOOL := FALSE; // 故障标志（非有限入参）[-] / the fault flag, a non finite input
END_VAR
VAR CONSTANT
    DL_QUA_EPS : LREAL := 1.0E-12; // 系数与判别式零阈值 [无量纲] / the coefficient and discriminant zero threshold
END_VAR
VAR
    lrD  : LREAL; // 判别式工作量 [无量纲] / the discriminant work value
    lrS  : LREAL; // 判别式平方根工作量 [无量纲] / the discriminant square root work value
    lrT  : LREAL; // 两倍二次项工作量 [无量纲] / the twice a work value
END_VAR

// 段 1｜返回值与输出预置安全值（四段式第一段，R45）/ segment 1, preset the return and the outputs
FC_DL_QuadraticSolve := FALSE; // 受理标志预置假 / preset the accepted flag false
fX1 := 0.0; // 根一预置零 / preset the root one zero
fX2 := 0.0; // 根二预置零 / preset the root two zero
nRoots := 0; // 根数预置零 / preset the count zero
bLinear := FALSE; // 线性标志预置假 / preset the linear flag false
bValid := FALSE; // 有效预置假 / preset the valid false
bError := FALSE; // 故障预置假 / preset the fault false

// 段 2｜非有限入参闸（三参数自反双判据全覆盖，R79）/ segment 2, the non finite gate
IF (fA <> fA) OR ((fA - fA) <> (fA - fA)) THEN // 二次项非有限 / a non finite a
    bError := TRUE; // 置故障 / raise the fault
END_IF
IF (fB <> fB) OR ((fB - fB) <> (fB - fB)) THEN // 一次项非有限 / a non finite b
    bError := TRUE; // 置故障 / raise the fault
END_IF
IF (fC <> fC) OR ((fC - fC) <> (fC - fC)) THEN // 常数项非有限 / a non finite c
    bError := TRUE; // 置故障 / raise the fault
END_IF
IF bError THEN // 非有限命中早退 / a non finite hit, return early
    RETURN; // 早退 / return early
END_IF

// 段 3｜a ≈ 0 退化线性分支（ABS 阈值禁等号，除零前置闸）/ segment 3, the degenerate linear branch
IF ABS(fA) < DL_QUA_EPS THEN // 二次项近似零 / the a near zero
    bLinear := TRUE; // 线性分支受理 / accept the linear branch
    IF ABS(fB) < DL_QUA_EPS THEN // 一次项也近似零 / the b near zero too
        IF ABS(fC) < DL_QUA_EPS THEN // 常数项也近似零：恒成立 / the c near zero too, an identity
            nRoots := -1; // 全 x 均为解（信息级）/ every x is a root, informational
        ELSE // 常数项非零：无解 / a nonzero c, no solution
            nRoots := 0; // 无实根（信息级非故障）/ no real root, informational
        END_IF
    ELSE // 正常线性 bx + c = 0 / the normal linear form
        nRoots := 1; // 单实根 / one real root
        fX1 := -fC / fB; // 求根（|fB| ≥ eps 已由分支保证，除零闸）/ the root, divided by the gated b
    END_IF
    bValid := TRUE; // 结果可用 / the result usable
    FC_DL_QuadraticSolve := TRUE; // 受理 / accept
    RETURN; // 早退（线性分支完结）/ return early
END_IF

// 段 4｜判别式三域分档（D ≥ 0 才开方，除 2a 前显式闸，边界二三）/ segment 4, the discriminant three domains
lrD := (fB * fB) - (4.0 * fA * fC); // 判别式 / the discriminant
IF lrD > DL_QUA_EPS THEN // 两实根域 / the two roots domain
    lrS := SQRT(lrD); // 开方（D > eps 已闸）/ the square root, gated
    lrT := 2.0 * fA; // 两倍二次项 / the twice a
    IF ABS(lrT) < DL_QUA_EPS THEN // 除零兜底闸（与段 3 判据互斥，防御纵深）/ the divide by zero fallback gate
        bError := TRUE; // 置故障 / raise the fault
        RETURN; // 早退 / return early
    END_IF
    fX1 := (-fB + lrS) / lrT; // 根一（公式分子取加号）/ the root one
    fX2 := (-fB - lrS) / lrT; // 根二 / the root two
    IF fX1 < fX2 THEN // 排序保证 x1 ≥ x2 / sort to keep x1 the larger
        fX1 := fX2; // 大根归 x1 / the larger to x1
        fX2 := (-fB + lrS) / lrT; // 小根归 x2 / the smaller to x2
    END_IF
    nRoots := 2; // 两实根 / two real roots
ELSIF lrD < -DL_QUA_EPS THEN // 无实根域（信息级非故障）/ the no real root domain
    nRoots := 0; // 无实根 / no real root
ELSE // 重根域 |D| ≤ eps / the double root domain
    lrT := 2.0 * fA; // 两倍二次项 / the twice a
    IF ABS(lrT) < DL_QUA_EPS THEN // 除零兜底闸 / the divide by zero fallback gate
        bError := TRUE; // 置故障 / raise the fault
        RETURN; // 早退 / return early
    END_IF
    fX1 := -fB / lrT; // 重根 x1 = x2 / the double root
    fX2 := fX1; // 重根同值 / the same value
    nRoots := 1; // 单重根 / one double root
END_IF
bValid := TRUE; // 结果可用 / the result usable
FC_DL_QuadraticSolve := TRUE; // 受理 / accept
END_FUNCTION

(* ---- FC_DL_QuantileCalc.st ---- *)
(*
  FC_DL_QuantileCalc  —  排序数组分位数（线性插值法） / Quantile of a sorted array by linear interpolation
  分类 Category : DL_MathData
  版本 Version  : 1.0.0
  来源 Source   : t2-1-lgf-math — 统计底座族零检索深化（P50/P95 工艺窗）
  溯源 Origin   : clean-room 实现，未复制任何源码行
  功能 Function : 1) 对前 nCnt 个已升序元素计算分位数 fQ，落位索引 pos := (nCnt-1) × fQ；
                  2) 正好整除点（pos 与 TRUNC(pos) 差 < 1.0E-9）直接取位，置信息级 04A6；
                  3) 非整除点在相邻两元素间线性插值；
                  4) fQ 越界按 [0, 1] 钳位并置信息级 04A5（钳位后照常输出）。
  边界 Boundary : ① 判界先行：nCnt <= 0 或 > 32 → 故障级 03E2，直接出口；
                  ② 样本非有限（NaN 自反判 / Inf 差值自减判）→ 故障级 03E3，拒绝输出；
                  ③ 整除点判定禁浮点 = 判等，用容差 1.0E-9；
                  ④ 无 GVL 依赖：纯函数，无外部变量引用，无物理 IO 地址。
  依赖 Depends  : 仅 Standard.library（TRUNC / ABS / LREAL 算术）
  码表 Error codes（段 0001，窗口 03E2~03E3 / 04A5~04A6）:
    16#0001_03E2 故障级：入参非法（nCnt <= 0 或 > 32），返回 0，bValid = FALSE，bError = TRUE
    16#0001_03E3 故障级：参与样本含非有限元素，返回 0，bValid = FALSE，bError = TRUE
    16#0001_04A5 信息级：fQ 越界已钳位至 [0, 1]（结果照常输出）
    16#0001_04A6 信息级：整除点直接取位（未插值）
  修订历史 Revision :
    2026-11-19  v1.0.0  R41 首版（批次 1 · 序号 5）
*)

FUNCTION FC_DL_QuantileCalc : LREAL
VAR_INPUT
    aSorted     : ARRAY[1..32] OF LREAL;   // 已升序样本数组 [EU]，前 nCnt 个参与 / Sorted samples, first nCnt used
    nCnt        : INT;               // 参与元素数 [个]，域 1..32 / Element count, 1..32
    fQ          : REAL;              // 分位数 [无量纲]，域 [0,1]，越界钳位 / Quantile, clamped to 0..1
END_VAR
VAR_OUTPUT
    eErr        : UDINT;             // 事件码，0 = 正常 / Event code
    bError      : BOOL;              // 故障级标志 / Fault-level flag
    bValid      : BOOL;              // 返回值是否可用 / Result usable flag
END_VAR
VAR
    fQc         : LREAL;             // 钳位后的分位数（LREAL 口径）/ Clamped quantile
    fPos        : LREAL;             // 落位索引 [索引] / Floating position index
    fLo         : LREAL;             // 落位整数部分 [索引] / Integer part of the position
    nLo         : INT;               // 下位索引（1 基）/ Lower index, one based
    nHi         : INT;               // 上位索引（1 基）/ Upper index, one based
    fFrac       : LREAL;             // 落位小数部分 [无量纲] / Fractional part
    i           : INT;               // 非有限扫描游标 [索引] / Scan cursor
    bClamped    : BOOL;              // 钳位发生标志 / Clamped flag
END_VAR
VAR CONSTANT
    DL_QTC_N_MAX      : INT := 32;               // 数组容量上限 [个] / Array capacity bound
    DL_QTC_TOL_IDX    : LREAL := 1.0E-9;         // 整除点判定容差 [索引] / Integer-point tolerance
    DL_QTC_ERR_IN     : UDINT := 16#0001_03E2;   // 故障级：nCnt 界外 / Fault: count out of range
    DL_QTC_ERR_NAN    : UDINT := 16#0001_03E3;   // 故障级：样本非有限 / Fault: non-finite sample
    DL_QTC_INFO_CLAMP : UDINT := 16#0001_04A5;   // 信息级：fQ 已钳位 / Info: quantile clamped
    DL_QTC_INFO_EXACT : UDINT := 16#0001_04A6;   // 信息级：整除点取位 / Info: exact index hit
END_VAR

(* —— 段 1｜返回值与错误状态预置 —— *)
FC_DL_QuantileCalc := 0.0;          // 缺省返回 0 / default return zero
eErr := 16#0000_0000;               // 预置无事件 / preset no event
bError := FALSE;                    // 预置无故障 / preset no fault
bValid := FALSE;                    // 预置不可用 / preset unusable
bClamped := FALSE;                  // 钳位标志清零 / clear clamp flag

(* —— 段 2｜判界先行：nCnt 域闸 —— *)
IF (nCnt <= 0) OR (nCnt > DL_QTC_N_MAX) THEN
    eErr := DL_QTC_ERR_IN;          // 故障级：nCnt 界外
    bError := TRUE;                 // 故障码配对置位（R101）
    bValid := FALSE;                // 结果不可用
    RETURN;                         // 直接出口 / early exit
END_IF

(* —— 段 3｜样本非有限闸：NaN 自反判 + Inf 差值自减判，逐元素扫描 —— *)
FOR i := 1 TO nCnt DO
    IF (aSorted[i] <> aSorted[i]) OR ((aSorted[i] - aSorted[i]) <> (aSorted[i] - aSorted[i])) THEN
        eErr := DL_QTC_ERR_NAN;     // 故障级：样本非有限
        bError := TRUE;             // 故障码配对置位（R101）
        bValid := FALSE;            // 结果不可用
        RETURN;                     // 直接出口 / early exit
    END_IF
END_FOR

(* —— 段 4｜fQ 钳位（越界不拒，钳位后照常输出 + 信息级） —— *)
fQc := LREAL(fQ);                   // REAL 升位到 LREAL 口径 / widen to LREAL
IF fQc < 0.0 THEN
    fQc := 0.0;                     // 下界钳位 / clamp low
    bClamped := TRUE;               // 钳位标志
ELSIF fQc > 1.0 THEN
    fQc := 1.0;                     // 上界钳位 / clamp high
    bClamped := TRUE;               // 钳位标志
END_IF

(* —— 段 5｜落位与插值：pos := (nCnt-1) × fQ，整除点直接取位（进位点） —— *)
fPos := INT_TO_LREAL(nCnt - 1) * fQc;   // 浮点落位 / floating position
fLo := TRUNC(fPos);                     // 整数部分 / integer part
nLo := LREAL_TO_INT(fLo) + 1;           // 1 基下位索引 / one-based lower index
fFrac := fPos - fLo;                    // 小数部分 / fractional part
IF fFrac < DL_QTC_TOL_IDX THEN
    FC_DL_QuantileCalc := aSorted[nLo]; // 整除点：直接取位（禁浮点 = 判等）/ exact hit
    eErr := DL_QTC_INFO_EXACT;          // 信息级：整除点取位 / info level
ELSIF nLo >= nCnt THEN
    FC_DL_QuantileCalc := aSorted[nCnt];    // 上边界防御：小数溢出取末位 / upper boundary defense
ELSE
    nHi := nLo + 1;                     // 上位索引 / upper index
    FC_DL_QuantileCalc := aSorted[nLo] + (aSorted[nHi] - aSorted[nLo]) * fFrac;
                                        // 线性插值 / linear interpolation
END_IF

(* —— 段 6｜出口 —— *)
IF bClamped THEN
    eErr := DL_QTC_INFO_CLAMP;      // 信息级：钳位提示（覆盖整除点信息级，钳位优先报告）/ info level
END_IF
bValid := TRUE;                     // 结果可用 / result usable
END_FUNCTION

(* ---- FC_DL_QuantizeStep.st ---- *)
(*
    组件名称 : FC_DL_QuantizeStep
    所属子库 : DL_MathData
    当前版本 : 1.0.0
    兼 容 性 : CODESYS V3.5+ / TwinCAT 3 / 汇川 InoProShop；仅依赖 Standard.library
    功能描述 : 按非整数步距量化，把任意给定值对齐到 n × step（编码器分辨率、给定值网格、成本最小单位的通用内核）。
              取舍 ①：禁用平台 ROUND —— 三家平台的 ROUND 在 .5 上是「银行家舍入」还是「远离零」并不一致，
              本件一律 TRUNC(fQ + 0.5)：加法把半值抬到整数侧，TRUNC 再向零截，等价于「半值向正方向」，
              负值同样成立（TRUNC(-1.8) = -1），语义单一且可复现。
              取舍 ②：商超精确域（> 1E15）时按输入直通而不硬算 —— LREAL 尾数只有 53 位，
              此域内 step 已小于末位权重，量化结果与输入仅差舍入噪声，硬算只会输出一个看着精确的假值。
              取舍 ③：步距非法时返回输入本身而非 0 —— 量化是「修饰」而非「求值」，步距坏了就把原值放行，
              静默置 0 会把一个传感器读数变成零位，比报错危险得多。
    开源溯源 : 原创实现。与存量 FC_DL_RoundSat / FC_DL_TruncEx 的职责边界：那两件到「整数」，；本件为 IEC 61131-3 标准语义的道莅防御性实现（原创实现，零外部源码复制）。
              本件到「非整数步距」。无外部源码参考，码位与分级 100% 自有。
    本文件内含 : FUNCTION FC_DL_QuantizeStep（单 POU，无配套类型）
    依 赖 : 无 DL_ 内部依赖；Standard.library: 无
    红线自检 : R1 ✓ 零全局变量与外部变量 ｜ R2 ✓ 零物理 IO 地址
              R3 ✓ 纯 IEC 61131-3 ｜ R4 ✓ 步距闸 + 非有限闸 + 精确域闸 + 乘积溢出复检 + 残差容差判据
              R5 ✓ 全变量中英双语同行注释 ｜ R6 N/A 纯函数无顺序状态机，无 CASE 可写
              R7 N/A 无定时器、无沿检测实例 ｜ R8 ✓ 全部阈值与半步比例常量化
    错误码   : 16#0001_0438 [信息级] 商超精确域（> DL_QUANT_MAX_RATIO），按输入直通，bValid = TRUE
               16#0001_0439 [信息级] 残差越半步（浮点误差提示），不改结果，bValid = TRUE
               16#0001_0372 [故障级] 步距 ≤ DL_FLOAT_EPS，返回输入直通，bValid = FALSE
               16#0001_0373 [故障级] 输入非有限（NaN 或 ±INF），返回 0，bValid = FALSE
               16#0001_0374 [故障级] 量化结果超有限域已饱和，bValid = FALSE
    码位总账 : 16#0001_0438 用 / 16#0001_0439 用 ｜ 16#0001_0372 用 / 16#0001_0373 用 / 16#0001_0374 用
    遗留假设 : ① TRUNC 返回与入参同宽（LREAL），赋回 LREAL 变量无需显式转换 —— IEC 语义推导，未三平台实测。
              ② 商的溢出安全依赖「IEEE 754 除法溢出得 INF 而非陷阱」这一平台行为；若某平台开启 FPU 异常陷阱，
              需在任务配置中关闭后再用本件。此条为编译/运行门槛，未实测。
    修订历史 :
        2026-11-16  v1.0.0  首版，R21 批次 1 入库
*)
FUNCTION FC_DL_QuantizeStep : LREAL
VAR_INPUT
    fIn             : LREAL := 0.0;   // 待量化值，全域有限实数 [工程单位] / value to quantise, finite real in engineering units
    fStep           : LREAL := 1.0;   // 量化步距，必须 > 0，如 0.01 mm [工程单位] / quantisation step, must exceed zero [engineering unit]
    bRoundHalfUp    : BOOL := TRUE;   // TRUE = 四舍五入（半值向正方向）；FALSE = 向零截断 / TRUE rounds half up, FALSE truncates toward zero
END_VAR
VAR_OUTPUT
    eErr            : UDINT;          // 错误码，0=正常；16#0001_04XX 信息级 / 16#0001_03XX 故障级 / error id, 0=ok
    bError          : BOOL;           // 故障级标志，eErr 落 16#0001_03XX 时为 TRUE / fault flag, TRUE on fault-level eErr
    bValid          : BOOL;           // 返回值是否可用 / output valid flag
    fResidual       : LREAL;          // 量化残差 = 结果 − 输入，带符号 [工程单位] / residual, result minus input, signed [engineering unit]
END_VAR
VAR
    fQ              : LREAL;          // 商工作寄存器，量化前先转成「步距个数」[倍] / quotient register, the value expressed in steps [ratio]
    fRet            : LREAL;          // 量化结果 [工程单位] / quantised result [engineering unit]
    fQAbs           : LREAL;          // 商的绝对值，只用于精确域判据 [倍] / absolute quotient, used only by the exact domain test [ratio]
END_VAR
VAR CONSTANT
    DL_QUANT_MAX_RATIO  : LREAL := 1.0E15;                     // 商超此值即尾数无小数精度，量化无意义 [倍] / above this ratio the mantissa has no fractional resolution [ratio]
    DL_QUANT_HALF       : LREAL := 0.5;                        // 半步比例，四舍五入的抬升量 [无量纲] / half step lifting term for rounding [dimensionless]
    DL_FLOAT_EPS        : LREAL := 1.0E-12;                    // 浮点判等容差，残差越界判据用 [无量纲] / float tolerance used by the residual test [dimensionless]
    DL_LREAL_MAX_FINITE : LREAL := 1.7976931348623157E308;     // LREAL 最大有限值 [无量纲] / largest finite LREAL [dimensionless]
    DL_LREAL_ZERO       : LREAL := 0.0;                        // 零哨兵 [无量纲] / zero sentinel [dimensionless]
    DL_ERR_NONE         : UDINT := 16#0000_0000;               // 无故障 / no error
END_VAR

// 段 1｜返回值与错误状态预置 / segment 1, preset the return value and the error state
FC_DL_QuantizeStep := DL_LREAL_ZERO;    // 故障缺省返回 0 / fault default returns zero
eErr       := DL_ERR_NONE;              // 预置无错误 / preset no error
bError     := FALSE;                    // 预置无故障 / preset no fault
bValid     := FALSE;                    // 预置结果不可用 / preset unusable
fResidual  := DL_LREAL_ZERO;            // 预置残差 0 / preset the residual to zero

// 段 2｜步距闸：步距不可用时直通输入，绝不静默置 0 / segment 2, step gate, pass the input through instead of zeroing it
IF fStep <= DL_FLOAT_EPS THEN
    FC_DL_QuantizeStep := fIn;          // 原值直通（量化是修饰，不是求值）/ pass the raw value through
    eErr   := 16#0001_0372;             // 步距非法（故障级）/ illegal step, fault level
    bError := TRUE;                     // 置故障标志 / raise the fault flag
    RETURN;                             // bValid 保持 FALSE，调用方必须知情 / bValid stays FALSE, the caller must know
END_IF

// 段 3｜输入有限性闸 / segment 3, input finiteness gate
IF (fIn <> fIn) OR (ABS(fIn) > DL_LREAL_MAX_FINITE) THEN
    eErr   := 16#0001_0373;             // 输入非有限（故障级）/ non-finite input, fault level
    bError := TRUE;                     // 置故障标志 / raise the fault flag
    RETURN;                             // 返回 0，bValid 保持 FALSE / return zero, bValid stays FALSE
END_IF

// 段 4｜唯一一次求商，随后复用同一结果做精确域判据 / segment 4, one division reused by the exact domain test
fQ    := fIn / fStep;                   // 步距已过闸（> EPS），除零结构性不可能 / the step passed the gate, division by zero is structurally impossible
fQAbs := ABS(fQ);                       // 取幅值供判据 / magnitude for the test
IF fQAbs > DL_QUANT_MAX_RATIO THEN
    FC_DL_QuantizeStep := fIn;          // 精确域外按输入直通 / pass the input through outside the exact domain
    eErr   := 16#0001_0438;             // 商超精确域（信息级，不置 bError）/ quotient beyond the exact domain, info level
    bValid := TRUE;                     // 直通值可用 / the pass-through value is usable
    RETURN;                             // 带值返回 / return with the value
END_IF

// 段 5｜取整：只允许 TRUNC（禁平台 ROUND，银行家舍入三平台不一致）/ segment 5, integer snap with TRUNC only
IF bRoundHalfUp THEN
    fQ := fQ + DL_QUANT_HALF;           // 半值向正方向抬升，负值同样成立 / lifting the half step works for negative values as well
END_IF
fQ := TRUNC(fQ);                        // 向零截断，语义单一可复现 / truncation toward zero, single reproducible semantics

// 段 6｜回乘并复检溢出 / segment 6, multiply back and re-check the overflow
fRet := fQ * fStep;                     // 回到工程单位 / back to engineering units
IF ABS(fRet) >= DL_LREAL_MAX_FINITE THEN
    IF fRet > DL_LREAL_ZERO THEN
        fRet := DL_LREAL_MAX_FINITE;    // 正向饱和 / saturate positive
    ELSE
        fRet := -DL_LREAL_MAX_FINITE;   // 负向饱和 / saturate negative
    END_IF
    eErr   := 16#0001_0374;             // 结果溢出已饱和（故障级）/ result overflow saturated, fault level
    bError := TRUE;                     // 置故障标志 / raise the fault flag
END_IF

// 段 7｜残差与容差判据：越半步只提示，不改结果 / segment 7, residual test, hint only
fResidual := fRet - fIn;                                                        // 带符号残差 / signed residual
IF (ABS(fResidual) - fStep * DL_QUANT_HALF) > DL_FLOAT_EPS THEN
    IF eErr = DL_ERR_NONE THEN                                                  // 不覆盖已有更高优先级的码 / never overwrite a code already set
        eErr := 16#0001_0439;                                                   // 残差越半步（信息级，浮点误差提示）/ residual beyond half a step, info level
    END_IF
END_IF

// 段 8｜出口 / segment 8, exit
FC_DL_QuantizeStep := fRet;             // 输出量化结果 / publish the quantised result
bValid := NOT bError;                   // 故障态不可用，信息态可用 / unusable after a fault, usable after an info code
END_FUNCTION

(* ---- FC_DL_QuartileCalc.st ---- *)
// FC_DL_QuartileCalc v1.0.0
// 开源溯源：self-cleanroom / 统计族补口
(*
  道莅工业代码库 | DL_MathData | FC_DL_QuartileCalc
  版本: 1.0.0 | 日期: 2026-11-23 | 轮次: R75
  功能: 四分位数 Q1/Q2/Q3 计算（数据升序排序后线性插值口径：
        位置 p = 1 + k·(n-1)/4，k=1,2,3，相邻两元素加权）
  邻件关系: 与 PercentileLReal / PercentileRank（百分位单值/排名）同族 ——
            差异点：本件一次返回三值（Q1/Q2/Q3），口径为四分位专用，
            排序基准一致（升序），码位独立（16#0002_1D01）
  数组契约: aData 为显式上界 100 的定长数组，nCount 为有效元素数（1..100），
            超界元素忽略；内部复制工作副本，不改调用方数组
*)
FUNCTION FC_DL_QuartileCalc : BOOL
VAR_INPUT
    aData  : ARRAY[1..100] OF REAL;              // 输入数据（前 nCount 个有效）[工程单位] / Input data, first nCount valid
    nCount : INT;                                // 有效元素数 [个]，域 1..100 / Valid element count, domain 1..100
END_VAR
VAR_OUTPUT
    fQ1     : REAL;                              // 下四分位 Q1 [工程单位] / First quartile
    fQ2     : REAL;                              // 中位数 Q2 [工程单位] / Median
    fQ3     : REAL;                              // 上四分位 Q3 [工程单位] / Third quartile
    bValid  : BOOL;                              // 结果有效回执 [-] / Result validity receipt
    uErrorId: UDINT;                             // 事件码，0 = 无事件；16#0002_1D01 = 计数非法 / Event code
END_VAR
VAR
    aWork   : ARRAY[1..100] OF REAL;             // 排序工作副本 [工程单位] / Working copy for sorting
    n       : INT;                               // 生效元素数 [个] / Effective count
    i       : INT;                               // 冒泡外层索引 [次] / Bubble outer index
    j       : INT;                               // 冒泡内层索引 [次] / Bubble inner index
    fSwap   : REAL;                              // 交换暂存 [工程单位] / Swap temp
    fPos    : REAL;                              // 四分位实数位置 [1] / Quartile real position
    nLo     : INT;                               // 位置下邻索引 [1] / Position lower index
    nHi     : INT;                               // 位置上邻索引 [1] / Position upper index
    fFrac   : REAL;                              // 插值份额 ∈ [0,1] [1] / Interpolation fraction
END_VAR

// —— 段 0：全路径缺省 —— //
fQ1 := 0.0;                                      // Q1 缺省零 / Q1 default
fQ2 := 0.0;                                      // Q2 缺省零 / Q2 default
fQ3 := 0.0;                                      // Q3 缺省零 / Q3 default
bValid := FALSE;                                 // 有效回执预清 / Validity preset
uErrorId := 16#0000;                             // 事件码预清 / Event code preset
FC_DL_QuartileCalc := FALSE;                     // 返回值缺省 FALSE / Return default FALSE

// —— 段 1：计数域闸（下标判界，R4） —— //
IF (nCount < 1) OR (nCount > 100) THEN           // 计数越出 1..100 / Count out of bounds
    uErrorId := 16#0002_1D01;                    // 信息级：计数非法（不置 bError） / Info level: illegal count
    RETURN;                                      // 不计算返回 / Return without computation
END_IF
n := nCount;                                     // 生效计数 / Effective count

// —— 段 2：复制工作副本（防调用方数组被改序） —— //
FOR i := 1 TO n DO                                // 逐元素复制（下标 i ≤ n ≤ 100 判界安全）/ Copy elements, index safe
    aWork[i] := aData[i];
END_FOR

// —— 段 3：冒泡升序排序（n ≤ 100，O(n²) 可接受） —— //
FOR i := 1 TO (n - 1) DO                          // 外层趟数 / Outer passes
    FOR j := 1 TO (n - i) DO                      // 内层相邻比较 / Inner adjacent compares
        IF aWork[j] > aWork[j + 1] THEN           // 升序交换 / Ascending swap
            fSwap := aWork[j];
            aWork[j] := aWork[j + 1];
            aWork[j + 1] := fSwap;
        END_IF
    END_FOR
END_FOR

// —— 段 4：单元素特判（四分位退化全等于该值，防 nLo 越界） —— //
IF n = 1 THEN                                     // 单元素：Q1=Q2=Q3 / Single element: all quartiles equal
    fQ1 := aWork[1];
    fQ2 := aWork[1];
    fQ3 := aWork[1];
    bValid := TRUE;
    FC_DL_QuartileCalc := TRUE;
    RETURN;
END_IF

// —— 段 5：线性插值四分位（位置法 p = 1 + k(n-1)/4） —— //
FOR i := 1 TO 3 DO                                // k = 1..3 依次算 Q1/Q2/Q3 / k=1..3 for Q1/Q2/Q3
    fPos := 1.0 + DINT_TO_REAL(i) * DINT_TO_REAL(n - 1) / 4.0;   // 实数位置 [1] / Real position
    nLo := REAL_TO_DINT(fPos);                    // 向零截断取下邻 / Truncate to lower index
    IF DINT_TO_REAL(nLo) > fPos THEN              // 截断上偏修正（负值域防御）/ Truncation correction
        nLo := nLo - 1;
    END_IF
    IF nLo < 1 THEN
        nLo := 1;                                 // 下界钳位 / Clamp low
    END_IF
    IF nLo > (n - 1) THEN
        nLo := n - 1;                             // 上邻必存在的上界钳位 / Clamp so upper neighbor exists
    END_IF
    nHi := nLo + 1;                               // 上邻索引 ≤ n 判界安全 / Upper neighbor safe
    fFrac := fPos - DINT_TO_REAL(nLo);            // 插值份额 / Interpolation fraction
    IF fFrac < 0.0 THEN
        fFrac := 0.0;                             // 份额下钳 / Fraction clamp low
    END_IF
    IF fFrac > 1.0 THEN
        fFrac := 1.0;                             // 份额上钳 / Fraction clamp high
    END_IF
    IF i = 1 THEN
        fQ1 := aWork[nLo] + fFrac * (aWork[nHi] - aWork[nLo]);   // Q1 插值 / Q1 interpolation
    ELSIF i = 2 THEN
        fQ2 := aWork[nLo] + fFrac * (aWork[nHi] - aWork[nLo]);   // Q2 插值 / Q2 interpolation
    ELSE
        fQ3 := aWork[nLo] + fFrac * (aWork[nHi] - aWork[nLo]);   // Q3 插值 / Q3 interpolation
    END_IF
END_FOR
bValid := TRUE;                                   // 有效回执 / Validity receipt
FC_DL_QuartileCalc := TRUE;                       // 返回成功 / Return success
END_FUNCTION
